METHOD get_stTankLevel : ST_Tank_Level
VAR_INPUT
END_VAR
VAR
	blank: ST_Tank_Level;
END_VAR
IF __ISVALIDREF(stTankLevel) THEN;
	get_stTankLevel:=stTankLevel;
ELSE;
	get_stTankLevel:=blank;
END_IF
END_METHOD

METHOD get_stTankLevel_OverFlow : BOOL
VAR_INPUT
END_VAR
VAR
	blank: ST_Tank_Level;
END_VAR
IF __ISVALIDREF(stTankLevel) THEN;
	IF stTankLevel.bIn_HL_signal 
	OR stTankLevel.rTankLevelPercentage>100
	OR (NOT MAIN.bTemp_Water_Overweight_check)
	THEN;
		get_stTankLevel_OverFlow:=TRUE;
	ELSE;
		get_stTankLevel_OverFlow:=FALSE;
	END_IF	
ELSE;
	get_stTankLevel_OverFlow:=FALSE;
END_IF
END_METHOD

END_FUNCTION_BLOCK

// ---- 00 Library/04 Recipe/FB_Recipe.TcPOU
FUNCTION_BLOCK FB_Recipe
VAR_INPUT
	pstRecipe				:POINTER TO ST_Recipe;
	bMemoRecipeUpdated		:BOOL:=FALSE;
	sRecipeDef				:STRING; (* current recipe definition *)
	bLoadDefault			:BOOL;
	sRecipesStoragePath		:STRING;
	bHMI_FrameActive		:BOOL;

END_VAR

VAR
	i						:INT;	
	RecipeManCommands 		:RecipeManCommands; (* Recipe Manager *)
	k						:INT;
	t1						:TON;
	check					:DWORD;
	INDEX					:INT:= 0;
	bReloadRecipes			:BOOL;
	rt_LoadDefault: R_TRIG;
	MessageBox			:MessageBox_Struct;
	arrLastReturn		: ARRAY[0..15] OF DWORD;
	LastReturn			:  DWORD;
	ton_RecipeUpdated: TON;
	sMessage: STRING;
	ton_SetStoragePath_Delay: TON;
	bSetStoragePath: BOOL:=TRUE;
	ton_SetStoragePathTimeOut: TON;
	bReturn: BOOL;
	
	ton_MessClear: TON;
	rt_Init: R_TRIG;
	sLastMessage: STRING;
	rt_Saved: R_TRIG;
	rt_FrameAvtive: R_TRIG;
	rt_LoadDefault1: R_TRIG;
END_VAR

act_SetStoragePath();
act_Disp();

IF pstRecipe^.bValidSelected THEN
	pstRecipe^.sSelectedReceipe:= pstRecipe^.arrRecipeNames[pstRecipe^.iRecipeIndex];
	pstRecipe^.bValidSelected:=FALSE;
END_IF

rt_FrameAvtive(CLK:=bHMI_FrameActive);
rt_LoadDefault1(CLK:=bLoadDefault);
IF pstRecipe^.bReInit OR rt_LoadDefault1.Q OR rt_FrameAvtive.Q THEN;
	pstRecipe^.bReInit:=FALSE;
	pstRecipe^.bInit:=FALSE;
	bSetStoragePath:=TRUE;
END_IF

t1(IN:=NOT pstRecipe^.bInit , PT:=T#0.5S);
IF (NOT pstRecipe^.bInit AND t1.Q) THEN
	
	IF NOT bSetStoragePath THEN;
		arrLastReturn[3]:=RecipeManCommands.ResetLastInfo();
		arrLastReturn[4]:=RecipeManCommands.ReloadRecipes(RecipeDefinitionName:=sRecipeDef);
		pstRecipe^.iRecipeCount:=RecipeManCommands.GetRecipeCount(sRecipeDef);
		FOR i := 0 TO GVL_Recipe.C_Max_RecipeFileNum DO
			pstRecipe^.arrRecipeNames[i] := '';
		END_FOR
		FOR i := 0 TO 1200 DO
			pstRecipe^.arrVariableNamesValue[i] := '';
			pstRecipe^.arrVariableValue[i] := '';
		END_FOR	
		(* save all recipe names of one recipe definition in an array *)
		arrLastReturn[0]:=RecipeManCommands.GetRecipeNames(sRecipeDef, ADR(pstRecipe^.arrRecipeNames),GVL_Recipe.C_Max_RecipeFileNum, 0);
		pstRecipe^.iRecipeIndex:=0;
		pstRecipe^.sLastSelectedReceipe:=pstRecipe^.sSelectedReceipe:=pstRecipe^.arrRecipeNames[0];
		pstRecipe^.bInit:=TRUE;
		pstRecipe^.bReInit:=FALSE;		
	END_IF

END_IF


rt_Init(CLK:=pstRecipe^.bInit);
IF pstRecipe^.bInit THEN

	IF pstRecipe^.sSelectedReceipe <> pstRecipe^.sLastSelectedReceipe 
	OR rt_Init.Q 
	OR rt_Saved.Q
	THEN;
				 
		arrLastReturn[1]:=RecipeManCommands.GetRecipeValues
			(
			RecipeDefinitionName:= sRecipeDef,
			RecipeName:= pstRecipe^.sSelectedReceipe, 
			pStrings:= ADR(pstRecipe^.arrVariableValue), 
			iSize:= 1200, 
			iStartIndex:= 0, 
			iStringLength:=80
			 );		
					
		arrLastReturn[2]:=RecipeManCommands.GetRecipeVariableNames
			(
			RecipeDefinitionName:=sRecipeDef,
			RecipeName:=pstRecipe^.sSelectedReceipe, 
			pStrings:= ADR(pstRecipe^.arrVariableNamesValue), 
			iSize:= 1200, 
			iStartIndex:= 0
			);
				
			pstRecipe^.bShowFile:=FALSE;
	END_IF
	pstRecipe^.sLastSelectedReceipe:=pstRecipe^.sSelectedReceipe;
END_IF


FOR i:=0 TO 15 DO
	IF arrLastReturn[i]<>0 THEN
		LastReturn:=arrLastReturn[i];
		EXIT;
	END_IF
	IF i=15 AND arrLastReturn[i]=0 THEN
		LastReturn:=0;
	END_IF
END_FOR

act_Cmd_List();

ACTION act_Cmd_List:
rt_LoadDefault(CLK:=bLoadDefault AND NOT bSetStoragePath);
IF rt_LoadDefault.Q THEN;
	pstRecipe^.sSelectedReceipe:='Default';
	pstRecipe^.bWriteToPLC_Cmd:=TRUE;
END_IF


IF pstRecipe^.bReloadRecipes THEN
	arrLastReturn[3]:=RecipeManCommands.ResetLastInfo();
	arrLastReturn[4]:=RecipeManCommands.ReloadRecipes(RecipeDefinitionName:=sRecipeDef);
	pstRecipe^.bReloadRecipes:=FALSE;
END_IF


IF pstRecipe^.bGetLastError THEN
	arrLastReturn[5]:=RecipeManCommands.GetLastError();
	pstRecipe^.bGetLastError:=FALSE;
END_IF


IF pstRecipe^.bResetLastError THEN
	arrLastReturn[6]:=RecipeManCommands.ResetLastError();
	pstRecipe^.bResetLastError:=FALSE;
	sMessage:='';
	FOR i:=0 TO 15 DO
		arrLastReturn[i]:=0;
	END_FOR	
END_IF

rt_Saved(CLK:=NOT pstRecipe^.bSaveFileCmd);
IF pstRecipe^.bSaveFileCmd  THEN
	sMessage:='cmd Save Recipe';
	IF  METH_Search(pstRecipe:=pstRecipe , sSearchRecipe:=pstRecipe^.sSelectedReceipe ) THEN
		//arrLastReturn[7]:=RecipeManCommands.ReadAndSaveRecipeAs(RecipeDefinitionName:=sRecipeDef,
		arrLastReturn[7]:=RecipeManCommands.ReadAndSaveRecipe(RecipeDefinitionName:=sRecipeDef,
			RecipeName:=pstRecipe^.sSelectedReceipe);// ,
			//FileName:='.txtrecipe' );
		sMessage:='cmd Save Recipe - Done';
		pstRecipe^.bSaveFileCmd:=FALSE;
	ELSE;
		sMessage:='cmd Save Recipe - Failed';
	END_IF
END_IF


IF pstRecipe^.bWriteToPLC_Cmd  THEN
	sMessage:='cmd Load Recipe';
	bMemoRecipeUpdated:=FALSE;
	IF  METH_Search(pstRecipe:=pstRecipe , sSearchRecipe:=pstRecipe^.sSelectedReceipe ) THEN
		arrLastReturn[8]:=RecipeManCommands.LoadRecipe(RecipeDefinitionName:= sRecipeDef, RecipeName:= pstRecipe^.sSelectedReceipe);
		arrLastReturn[9]:=RecipeManCommands.WriteRecipe(RecipeDefinitionName:= sRecipeDef, RecipeName:= pstRecipe^.sSelectedReceipe);
		sMessage:='cmd Load Recipe - Done';
		pstRecipe^.bWriteToPLC_Cmd:=FALSE;
		ton_RecipeUpdated.IN:=TRUE;
	ELSE;
		sMessage:='cmd Load Recipe - Failed';
	END_IF
END_IF
ton_RecipeUpdated(PT:=T#1S);
IF ton_RecipeUpdated.Q THEN;
	bMemoRecipeUpdated:=TRUE;	
	ton_RecipeUpdated.IN:=FALSE;
END_IF


IF pstRecipe^.bCreateRecipe AND pstRecipe^.sNewRecipeName <> '' THEN
	arrLastReturn[10]:=RecipeManCommands.CreateRecipe(sRecipeDef ,pstRecipe^.sNewRecipeName);
	sMessage:='cmd Create Recipe - Done';
	pstRecipe^.bCreateRecipe:=FALSE;
	pstRecipe^.bReInit:=TRUE;
END_IF


IF pstRecipe^.bDeleteRecipe THEN
	sMessage:='cmd Delete Recipe';
	IF  METH_Search(pstRecipe:=pstRecipe , sSearchRecipe:=pstRecipe^.sSelectedReceipe ) THEN
		arrLastReturn[11]:=RecipeManCommands.DeleteRecipe(sRecipeDef ,pstRecipe^.sSelectedReceipe);
		sMessage:='cmd Delete Recipe - Done';
		pstRecipe^.bDeleteRecipe:=FALSE;
		pstRecipe^.bReInit:=TRUE;
	ELSE;
		sMessage:='cmd Delete Recipe - Failed';
	END_IF
END_IF

ton_MessClear(PT:=T#30S);
IF sMessage<>sLastMessage THEN;
	ton_MessClear(IN:=FALSE);
	sLastMessage:=sMessage;
ELSIF sMessage<>'' THEN;
	ton_MessClear.IN:=TRUE;
ELSE;
	ton_MessClear.IN:=FALSE;
END_IF
IF ton_MessClear.Q THEN;
	sMessage:='';
END_IF
END_ACTION

ACTION act_Disp:

IF pstRecipe^.iDispSel<0 THEN; pstRecipe^.iDispSel:=0; END_IF
IF pstRecipe^.iDispSel>1180 THEN; pstRecipe^.iDispSel:=1180; END_IF

//FOR k:=iDispSel TO iDispSel+19 DO;
FOR k:=0 TO 20 DO;
	pstRecipe^.arrVariableDisp[0,k]:= INT_TO_STRING(pstRecipe^.iDispSel+k);
	pstRecipe^.arrVariableDisp[1,k]:=pstRecipe^.arrVariableNamesValue[pstRecipe^.iDispSel+k];
	pstRecipe^.arrVariableDisp[2,k]:=pstRecipe^.arrVariableValue[pstRecipe^.iDispSel+k];
END_FOR
END_ACTION

ACTION act_SetStoragePath:
ton_SetStoragePath_Delay(PT:=T#0.5S,IN:=bSetStoragePath);
ton_SetStoragePathTimeOut(PT:=T#2S);

IF ton_SetStoragePath_Delay.Q THEN;
	bReturn:=RecipeManCommands.SetStoragePath(stPath:=sRecipesStoragePath);
	//sMessage:='cmd Set Storage Path';
	IF bReturn THEN;
		bSetStoragePath:=FALSE;
		ton_SetStoragePathTimeOut.IN:=FALSE;
		//sMessage:='cmd Set Storage Path - Done';
	ELSE
		ton_SetStoragePathTimeOut.IN:=TRUE;
	END_IF
	
	IF ton_SetStoragePathTimeOut.Q THEN;
		bSetStoragePath:=FALSE;
		ton_SetStoragePathTimeOut.IN:=FALSE;
		//sMessage:='cmd Set Storage Path - Failed';		
	END_IF
END_IF
END_ACTION

METHOD METH_Search : BOOL
VAR_INPUT
	pstRecipe :POINTER TO ST_Recipe;
	sSearchRecipe	:STRING(30);
END_VAR

VAR
	i: INT;
END_VAR
METH_Search:=FALSE;
FOR i:= 0 TO GVL_Recipe.C_Max_RecipeFileNum DO
	IF sSearchRecipe = pstRecipe^.arrRecipeNames[i] THEN
		METH_Search:=TRUE;
		EXIT;
	END_IF
END_FOR
END_METHOD

END_FUNCTION_BLOCK

// ---- 00 Library/04-Messages/FB_PrintErrMessageByID.TcPOU
FUNCTION_BLOCK FB_PrintErrMessageByID
VAR_INPUT
	sActErrorID			: STRING;
	iFB_Num				: INT:=0;
	sModuleDescription	:STRING:='';
END_VAR
VAR_OUTPUT
END_VAR
VAR
	cFound				: INT;
	i					: INT;
	iFound				: INT;
	bNewMeasege			: BOOL;
	rtrig1				: R_TRIG;
	sLastErrorID		: STRING;
	j: INT;
	sFB_Num: STRING(3);

END_VAR




	
	IF sActErrorID<>'000x000x000'  AND sActErrorID<>'' THEN
		IF iFB_Num>0 THEN;
			sFB_Num:=F_iFB_Num_sFB_Num(iFB_Num:=iFB_Num);
			sLastErrorID:=REPLACE(sActErrorID,sFB_Num,3,5);
		ELSE;
			sLastErrorID:=sActErrorID;
		END_IF			
		
		bNewMeasege:=TRUE;
		FOR i:=1 TO 100 DO
			IF Buffer_Act_Message[i].sErrID=sLastErrorID THEN;//sActErrorID
				//IF Buffer_Act_Message[i].sModuleDescription = sFB_ModuleDescription THEN
					bNewMeasege:=FALSE;
					EXIT; 
				//END_IF
			END_IF
		END_FOR
	ELSE
		bNewMeasege:=FALSE;
	END_IF
	
	IF bNewMeasege THEN;
		FOR i:=100 TO 2 BY -1 DO
			Buffer_Act_Message[i].sDateTime:=Buffer_Act_Message[i-1].sDateTime;
			Buffer_Act_Message[i].sErrID:=Buffer_Act_Message[i-1].sErrID;
			Buffer_Act_Message[i].sErrorMessage:=Buffer_Act_Message[i-1].sErrorMessage;
			Buffer_Act_Message[i].sLevel:=Buffer_Act_Message[i-1].sLevel;
			Buffer_Act_Message[i].sModuleDescription:=Buffer_Act_Message[i-1].sModuleDescription;
		END_FOR
		
		Buffer_Act_Message[1].sDateTime:=prg_RealClock.sRealTime_Date;
		Buffer_Act_Message[1].sErrID:=sLastErrorID;//sActErrorID
		Buffer_Act_Message[1].sModuleDescription:=sModuleDescription;

		//IF sActErrorID='000x000x999' THEN;
		//	Buffer_Act_Message[1].sErrorMessage:='General Error';	(*	Error description Not Found	*)
		//ELSE
			cFound:=0;
			FOR i:=1 TO C_Max_ErrorList DO
				IF ar_ErrorList[i,eErrID]=sActErrorID THEN
					iFound:=i;
					ar_ErrorActive[iFound]:=TRUE;
					cFound:=cFound+1;
				END_IF
			END_FOR
	
			IF cFound=1 THEN;
				Buffer_Act_Message[1].sErrorMessage:=ar_ErrorList[iFound,eErrMeassage];	(*	Error from the List	*)
				Buffer_Act_Message[1].sLevel:=ar_ErrorList[iFound,eErrLevel];	(*	Error Level from the List	*)
			ELSIF cFound=0 THEN; //(*	Error ID not Foud on the Error_List*)
				Buffer_Act_Message[1].sErrorMessage:='Error ID not found on the "Error_List"';	
				Buffer_Act_Message[1].sLevel:='Unknown';
			ELSIF cFound>1 THEN; //(*	More then one Errors Foud with the same  ID*)
				Buffer_Act_Message[1].sErrorMessage:='More then one error with the same ID  found on the "Error_list"';	
				Buffer_Act_Message[1].sLevel:='Unknown';
			END_IF
		//END_IF
		FUN_Write_Line_To_History();
	END_IF

END_FUNCTION_BLOCK

// ---- 00 Library/04-Messages/F_iFB_Num_sFB_Num.TcPOU
FUNCTION F_iFB_Num_sFB_Num : STRING(3)
VAR_INPUT
	iFB_Num: INT;
END_VAR
VAR
END_VAR

IF iFB_Num<10 THEN;
	F_iFB_Num_sFB_Num:=CONCAT(STR1:='00',STR2:=INT_TO_STRING(iFB_Num));
ELSIF iFB_Num<100 THEN;
	F_iFB_Num_sFB_Num:=CONCAT(STR1:='0',STR2:=INT_TO_STRING(iFB_Num));
ELSE;
	F_iFB_Num_sFB_Num:=CONCAT(STR1:='',STR2:=INT_TO_STRING(iFB_Num));
END_IF

END_FUNCTION

// ---- 00 Library/03 SFC/FB_SFC_Template.TcPOU
FUNCTION_BLOCK FB_SFC_Template EXTENDS FB_SFC_Cycle IMPLEMENTS ITF_FB_SFC_Cycle
VAR_INPUT
END_VAR
VAR_OUTPUT
END_VAR
VAR
END_VAR

m_Set_SFCFlags_Reference();
SUPER^();

ACTION act_Oper:
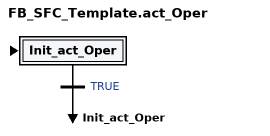
INITIAL_STEP Init_act_Oper:
END_STEP
TRANSITION FROM Init_act_Oper TO Init_act_Oper
    := TRUE;
END_TRANSITION
END_ACTION

METHOD m_Set_SFCFlags_Reference : BOOL
//Set reference to SFC flags

refSFC.SFCInit REF= SFCInit;
refSFC.SFCReset REF= SFCReset;
refSFC.SFCError REF= SFCError;
refSFC.SFCEnableLimit REF= SFCEnableLimit;
refSFC.SFCErrorStep REF= SFCErrorStep;
refSFC.SFCErrorPOU REF= SFCErrorPOU;
refSFC.SFCQuitError REF= SFCQuitError;
refSFC.SFCPause REF= SFCPause;
refSFC.SFCTrans REF= SFCTrans;
refSFC.SFCCurrentStep REF= SFCCurrentStep;
refSFC.SFCTip REF= SFCTip;
refSFC.SFCTipMode REF= SFCTipMode;

// Cycle handle for SFC
m_SFC_Handle();
END_METHOD

END_FUNCTION_BLOCK

// ---- 03 Project/00 -Initialise/prg_Initialise.TcPOU
PROGRAM prg_Initialise
VAR_INPUT
	ResumeSFC       : BOOL; 		(*	not automatic	*)
	//Added SFC Cycle handle Variables
	
	SFCInit             : BOOL;  //shachar
END_VAR

VAR


(* 8888888888888888   SFC   8888888888888888888888*)
	sCycleName	        : STRING;
	SFCCurrentStep      : STRING;
	SFCErrorPOU         : STRING;
	SFCErrorStep        : STRING;
	SFCError            : BOOL;
	SFCPause            : BOOL;
	
	SFCTipMode          : BOOL;
	SFCTip              : BOOL;
	SFCEnableLimit		: BOOL:=TRUE;
	// Reset Error
	SFCReset			: BOOL;
	ErrorSFC            : BOOL; 	(*	not automatic	*)

	ResetError          : BOOL; 	(*	not automatic	*)
	Last_SFCErrorStep   : STRING; 	(*	not automatic	*)
	//ErrorToPrint        : STRING; 	(*	not automatic	*)
	//Last_ErrorToPrint   : STRING; 	(*	not automatic	*)

 //   stSafety			:ST_BasicCycle;  //shachar
(* 8888888888888888   SFC   8888888888888888888888*)




	Pis             : INT;
	c_PisInitCheck  : INT;
	b_AllPisInitPos : BOOL;

	i               : INT;
	c_LatInitCheck  : INT;

	c_PisResetCleare: INT;

	k               : INT;

	bGeneralDone    : BOOL;
	bPistonDone     : BOOL;
	b_StationDone   : BOOL;
	bLoadConvDone   : BOOL;
	bUnloadConvDone : BOOL;
	bTableDone      : BOOL;
	bStackerDone    : BOOL;
    bManipulatorDone: BOOL;

	init_General    : BOOL;
	init_AllPiston  : BOOL;
	init_AllStation : BOOL;
	init_Table      : BOOL;
	init_LoadConv   : BOOL;
	init_UnloadConv : BOOL;
	init_Stacker    : BOOL;
	init_Manipulator: BOOL;

	bMessLoadInit   : BOOL;
	bMessUnloadInit : BOOL;
	
	sFB_ID          : STRING(4):='004';
	sFB_Num         : STRING(4):='000';
	sActErrorID     : STRING;
	//Added SFC Cycle handle Variables
	fb_SFC_Cycle		    : FB_SFC_Cycle;
	fbFormatString	    	: FB_FORMATSTRING;
	sFullErrorId		    : STRING(12);//sAAAxBBBxEEE
	bReset					: BOOL;

	bIntZoneOk: BOOL;
	bNotPrepare: BOOL;
	p_ManipReset: POINTER TO BOOL;
	p_PowerMotorOn: POINTER TO BOOL;
	p_SafetyStart: POINTER TO BOOL;
   // fbPowerMotorOn			:FB_PowerMotorOn;

	IndexOn: BOOL;
	LoadOn: BOOL;
	UnloadOn: BOOL;
	ManipOn: BOOL;
	p_PowerMotorPower: POINTER TO BOOL;
	p_PowerMotorOff: POINTER TO BOOL;
	iResumeCount: INT;
	iIndexCount: INT;
	iLoadCount: INT;
	iUnloadCount: INT;
	iManipCount: INT;
	p_ManipResume: POINTER TO BOOL;
END_VAR

VAR_IN_OUT
	stOperation	: ST_OperationButtons;	
END_VAR

act_General();
act_Piston();
act_GetErrorID();
fb_SFC_Cycle
( 
	sCycleName:= 'Initialize', 
	bSFCError:= SFCError, 
	sSFCCurrentStep:=SFCCurrentStep , 
	sSFCErrorStep:= SFCErrorStep, 
	sSFCErrorPOU:=SFCErrorPOU , 
	sActErrorID:=sFullErrorId,
	sFB_ModuleDescription:= fb_SFC_Cycle.sCycleName, 
	sLast_SFCErrorStep=>Last_SFCErrorStep , 
	bErrorSFC_Occured=> ErrorSFC, 
	//sErrorToPrint=>ErrorToPrint , 
	//sLast_ErrorToPrint=>Last_ErrorToPrint,
    bSFCInit=>SFCInit , 
	stOperation:= stOperation,
	bResumeSFC:=ResumeSFC , 
	bResetError:=ResetError , 
	bSFCPause:= SFCPause, 
	bResetCycle:=SFCReset
);



IF NOT bStateSafe	
OR init_AllPiston
THEN;
	bGeneralDone:=FALSE;
	bPistonDone:=FALSE;
	b_StationDone:=FALSE;
	bLoadConvDone:=FALSE;
	bUnloadConvDone:=FALSE;
	bTableDone:=FALSE;
	bStackerDone:=FALSE;
	bManipulatorDone:=FALSE;  //shachar
END_IF

ACTION act_General:
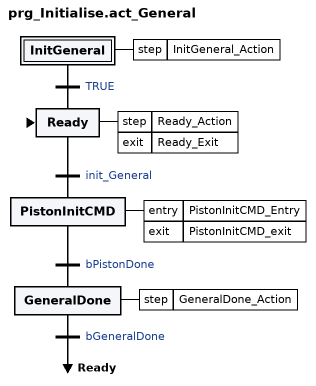
INITIAL_STEP InitGeneral:
    InitGeneral_Action(N);  // step action
END_STEP
TRANSITION FROM InitGeneral TO Ready
    := TRUE;
END_TRANSITION
STEP Ready:
    Ready_Action(N);  // step action
    Ready_Exit(P0);  // exit action
END_STEP
TRANSITION FROM Ready TO PistonInitCMD
    := init_General;
END_TRANSITION
STEP PistonInitCMD:  // min time t#2s
    PistonInitCMD_Entry(P1);  // entry action
    PistonInitCMD_exit(P0);  // exit action
END_STEP
TRANSITION FROM PistonInitCMD TO GeneralDone
    := bPistonDone;
END_TRANSITION
STEP GeneralDone:
    GeneralDone_Action(N);  // step action
END_STEP
TRANSITION FROM GeneralDone TO Ready
    := bGeneralDone;
END_TRANSITION
END_ACTION

ACTION act_GetErrorID:
IF ErrorSFC THEN;
	// Initialization
	IF    Last_SFCErrorStep='WatingForEmergencyOK' 			THEN sActErrorID:='001';
	ELSIF Last_SFCErrorStep='WatingForInterlockOK' 		    THEN sActErrorID:='002';
	ELSIF Last_SFCErrorStep='WatingForMotorsOK' 			THEN sActErrorID:='003';
	ELSIF Last_SFCErrorStep='CheckInitStationDone' 			THEN sActErrorID:='004';
	ELSIF Last_SFCErrorStep='Station_Initialization' 		THEN sActErrorID:='005';
	ELSIF Last_SFCErrorStep='Loader_Initialization' 		THEN sActErrorID:='006';
	ELSIF Last_SFCErrorStep='Unload_Station' 			    THEN sActErrorID:='007';
	ELSIF Last_SFCErrorStep='Measuring_Station' 			THEN sActErrorID:='008';
	ELSIF Last_SFCErrorStep='Gripper_Oriantation' 			THEN sActErrorID:='009';
	ELSIF Last_SFCErrorStep='Index_Homming' 			    THEN sActErrorID:='010';
	ELSIF Last_SFCErrorStep='PaletBypasCheck_1' 			THEN sActErrorID:='011';
	ELSIF Last_SFCErrorStep='PaletCheck_1' 			        THEN sActErrorID:='012';
	ELSIF Last_SFCErrorStep='Cover_Station' 			    THEN sActErrorID:='023';	
	ELSE;
		 sActErrorID:='999';
	END_IF
//ELSIF bWarning THEN;
	// Leave the warning message to print
ELSE;
		 sActErrorID:='000';
END_IF
//*** Error Format ***
fbFormatString(
	sFormat:= '%.3sx%.3sx%.3s', 
	arg1:= F_STRINGEx(sFB_ID), 
	arg2:= F_STRINGEx(sFB_Num), 
	arg3:= F_STRINGEx(sActErrorID), 
	sOut=>sFullErrorId );
	
//(*Clean Last ErrID*)IF NOT SFCPause THEN	sFullErrorId:='';END_IF
END_ACTION

ACTION act_Piston:
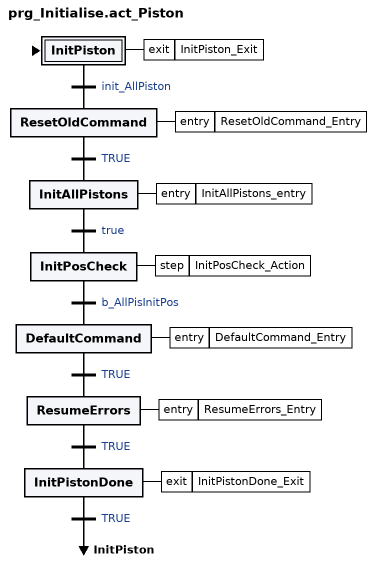
INITIAL_STEP InitPiston:
    InitPiston_Exit(P0);  // exit action
END_STEP
TRANSITION FROM InitPiston TO ResetOldCommand
    := init_AllPiston;
END_TRANSITION
STEP ResetOldCommand:  // min time T#0.1S
    ResetOldCommand_Entry(P1);  // entry action
END_STEP
TRANSITION FROM ResetOldCommand TO InitAllPistons
    := TRUE;
END_TRANSITION
STEP InitAllPistons:  // min time t#1s
    InitAllPistons_entry(P1);  // entry action
END_STEP
TRANSITION FROM InitAllPistons TO InitPosCheck
    := true;
END_TRANSITION
STEP InitPosCheck:
    InitPosCheck_Action(N);  // step action
END_STEP
TRANSITION FROM InitPosCheck TO DefaultCommand
    := b_AllPisInitPos;
END_TRANSITION
STEP DefaultCommand:  // min time T#0.2S
    DefaultCommand_Entry(P1);  // entry action
END_STEP
TRANSITION FROM DefaultCommand TO ResumeErrors
    := TRUE;
END_TRANSITION
STEP ResumeErrors:  // min time T#0.2S
    ResumeErrors_Entry(P1);  // entry action
END_STEP
TRANSITION FROM ResumeErrors TO InitPistonDone
    := TRUE;
END_TRANSITION
STEP InitPistonDone:
    InitPistonDone_Exit(P0);  // exit action
END_STEP
TRANSITION FROM InitPistonDone TO InitPiston
    := TRUE;
END_TRANSITION
END_ACTION

ACTION DefaultCommand_Entry:
	(*FOR Pis:=1 TO 24 BY 1 DO
		db_Lat[Pis].req_DefaultPos:=TRUE;
	END_FOR*)
	
	FOR Pis:=1 TO C_Max_Pistons BY 1 DO
		IF stPis[Pis].b_PistonActive THEN;
			stPis[Pis].req_Init:=TRUE;
		END_IF		
	END_FOR
END_ACTION

ACTION GeneralDone_Action:
init_General:=FALSE;
bGeneralDone:=TRUE;
END_ACTION

ACTION InitAllPistons_entry:
prg_Pistons.bInitAllPiston:=TRUE;
END_ACTION

ACTION InitGeneral_Action:
SFCReset:=FALSE;

init_AllPiston   :=FALSE;
END_ACTION

ACTION InitPiston_Exit:
	b_AllPisInitPos:=FALSE;
	bPistonDone:=FALSE;
END_ACTION

ACTION InitPistonDone_Exit:
	init_AllPiston:=FALSE;
	bPistonDone:=TRUE;
END_ACTION

ACTION InitPosCheck_Action:
			c_PisInitCheck:=0;
	FOR Pis:=1 TO C_Max_Pistons BY 1 DO
		IF fb_Pis[Pis].SFCCurrentStep<>'Ready' AND fb_Pis[Pis].SFCCurrentStep<>''THEN
			c_PisInitCheck:=c_PisInitCheck+1;
		END_IF
	END_FOR

			c_PisResetCleare:=0;
	FOR Pis:=1 TO C_Max_Pistons BY 1 DO
		IF stPis[Pis].b_Reset THEN
			c_PisResetCleare:=c_PisResetCleare+1;
		END_IF
	END_FOR

	(*		c_LatInitCheck:=0;
	FOR Pis:=1 TO 24 BY 1 DO
		IF fb_Lat[Pis].SFCCurrentStep<>'Ready' AND fb_Lat[Pis].SFCCurrentStep<>'' THEN
			c_LatInitCheck:=c_LatInitCheck+1;
		END_IF
	END_FOR*)


		IF 	c_PisInitCheck=0  AND c_LatInitCheck=0 (*AND 	c_PisResetCleare=0*) THEN
			b_AllPisInitPos:=TRUE;
		ELSE
			b_AllPisInitPos:=FALSE;
		END_IF
END_ACTION

ACTION PistonInitCMD_Entry:
init_AllPiston:=TRUE;
END_ACTION

ACTION PistonInitCMD_exit:
Global_Variables.ResumeAll :=TRUE;
END_ACTION

ACTION Ready_Action:
IF TRUE
AND	bPistonDone
(*AND	b_StationDone
AND	bLoadConvDone
AND	bUnloadConvDone
AND	bTableDone
AND (bManipulatorDone OR NOT b_ManipulatorExist)
AND	(bStackerDone OR NOT b_StackerExist)*)
THEN
	bGeneralDone:=TRUE;

ELSE
	bGeneralDone:=FALSE;
END_IF
END_ACTION

ACTION Ready_Exit:
bGeneralDone:=FALSE;
bPistonDone:=FALSE;
b_StationDone:=FALSE;
bLoadConvDone:=FALSE;
bUnloadConvDone:=FALSE;
bTableDone:=FALSE;
bStackerDone:=FALSE;

bManipulatorDone:=FALSE; //shachar
iResumeCount:=0;
END_ACTION

ACTION ResetOldCommand_Entry:
	(*FOR Pis:=1 TO 24 BY 1 DO
		db_Lat[Pis].req_Reset:=TRUE;
	END_FOR*)
	FOR Pis:=1 TO C_Max_Pistons BY 1 DO
		stPis[Pis].b_Reset:=TRUE;
	END_FOR
END_ACTION

ACTION ResumeErrors_Entry:
	(*FOR Pis:=1 TO 24 BY 1 DO
		db_Lat[Pis].req_Resume:=TRUE;
	END_FOR*)
	FOR Pis:=1 TO C_Max_Pistons BY 1 DO
		stPis[Pis].b_Resume:=TRUE;
	END_FOR
END_ACTION

END_PROGRAM

// ---- 03 Project/31 AnybusCommunication/FB_Anybus_Interface.TcPOU
//CIP <-> Siemens exchange through the Anybus Communicator, 128 bytes each direction.
//Spec: "Интерфейс CIP ↔ Siemens через Anybus", meeting 28.10.2026.
//Decodes the Siemens data, checks ALIVE and the values, encodes the CIP status.
//While communication is lost all Siemens inputs are treated as 0 (REQUEST ON drops -> CIP pause).
FUNCTION_BLOCK FB_Anybus_Interface
VAR_INPUT
	stStatus		: ST_Anybus_Outputs;	//CIP -> Siemens, filled by the CIP logic (bAlive is generated here)
	bFieldbusOk		: BOOL := TRUE;			//gateway EtherCAT slave: WcState = 0 (gIO.Anybus_WcState in MAIN)
	bSwapBytes		: BOOL := TRUE;			//TRUE: INT/DINT are big-endian (Profinet), swapped here
	tAliveTimeout	: TIME := T#2S;			//Siemens ALIVE must toggle within this time
	tNextStable		: TIME := T#3S;			//NEXT CLIENT / NEXT RECIPE must be stable this long
END_VAR
VAR_IN_OUT
	arRawIn			: ARRAY[0..127] OF BYTE;	//gIO.Anybus_Inputs_Raw
	arRawOut		: ARRAY[0..127] OF BYTE;	//gIO.Anybus_Outputs_Raw
END_VAR
VAR_OUTPUT
	stIn			: ST_Anybus_Inputs;		//Siemens -> CIP, all 0 while communication is lost
	stOut			: ST_Anybus_Outputs;	//CIP -> Siemens as actually sent (with ALIVE, alarm bit and code)
	bCommOk			: BOOL;					//fieldbus OK and Siemens ALIVE toggles
	eRequest		: E_Anybus_Request;		//combination of REQUEST ON / REQUEST OFF
	bRequestOnEdge	: BOOL;					//one cycle when eRequest becomes eOn (start or resume)
	bRequestOffEdge	: BOOL;					//one cycle when eRequest becomes eOff
	bCurrentValid	: BOOL;					//CLIENT ID, RECIPE TYPE, CLIENT TYPE are in range
	bNextValid		: BOOL;					//next client is in range and stable for tNextStable
	nNextClient		: INT;					//accepted next client, 0 = none
	eNextRecipe		: E_Anybus_RecipeType;	//accepted next recipe
	eNextClientType	: E_Anybus_ClientType;	//accepted next client type, eNone = not sent
	eAlarm			: E_Anybus_Alarm;		//interface alarm, eNone = OK
END_VAR
VAR
	stRaw			: ST_Anybus_Inputs;		//decoded, before the communication check
	stBlank			: ST_Anybus_Inputs;

	//ALIVE
	bAliveOut		: BOOL;
	tonAliveOut		: TON;
	tonAliveIn		: TON;
	bAliveInMemo	: BOOL;
	bAliveSeen		: BOOL;					//at least one toggle since start

	rtRequestOn		: R_TRIG;
	rtRequestOff	: R_TRIG;

	//Next client
	tonNextStable	: TON;
	nNextClientMemo	: INT;
	eNextRecipeMemo	: E_Anybus_RecipeType;
	eNextTypeMemo	: E_Anybus_ClientType;
	bNextInRange	: BOOL;
END_VAR
VAR CONSTANT
	cnClientMax		: INT := 30;
END_VAR

//Decode Siemens -> CIP
//Bits are addressed by byte (Siemens x.y = byte x, bit y), no swap
stRaw.bAlarm			:= arRawIn[0].0;
stRaw.bReady			:= arRawIn[0].1;
stRaw.bRequestOn		:= arRawIn[0].2;
stRaw.bRequestOff		:= arRawIn[0].3;
stRaw.bInletPumpEnable	:= arRawIn[0].4;
stRaw.bPause			:= arRawIn[0].5;
stRaw.bClientEmpty		:= arRawIn[0].6;
stRaw.bAlive			:= arRawIn[0].7;
stRaw.bSprinklerState	:= arRawIn[1].0;
stRaw.nClientId			:= m_GetInt(arRaw:=arRawIn, nWord:=1);
stRaw.eRecipeType		:= m_GetInt(arRaw:=arRawIn, nWord:=2);
stRaw.eClientType		:= m_GetInt(arRaw:=arRawIn, nWord:=3);
stRaw.nNextClient		:= m_GetInt(arRaw:=arRawIn, nWord:=4);
stRaw.eNextRecipe		:= m_GetInt(arRaw:=arRawIn, nWord:=5);
stRaw.eNextClientType	:= m_GetInt(arRaw:=arRawIn, nWord:=6);

//Siemens ALIVE watchdog
IF stRaw.bAlive <> bAliveInMemo THEN;
	bAliveInMemo:=stRaw.bAlive;
	bAliveSeen:=TRUE;
	tonAliveIn(IN:=FALSE);
END_IF
tonAliveIn(IN:=TRUE, PT:=tAliveTimeout);
bCommOk:=bFieldbusOk AND bAliveSeen AND NOT tonAliveIn.Q;

//Communication lost: the same as the gateway clearing the data
IF bCommOk THEN;
	stIn:=stRaw;
ELSE;
	stIn:=stBlank;
END_IF

//REQUEST ON / REQUEST OFF
IF stIn.bRequestOn AND stIn.bRequestOff THEN;
	eRequest:=E_Anybus_Request.eConflict;
ELSIF stIn.bRequestOn THEN;
	eRequest:=E_Anybus_Request.eOn;
ELSIF stIn.bRequestOff THEN;
	eRequest:=E_Anybus_Request.eOff;
ELSE;
	eRequest:=E_Anybus_Request.eNone;
END_IF
rtRequestOn(CLK:=eRequest=E_Anybus_Request.eOn);
bRequestOnEdge:=rtRequestOn.Q;
rtRequestOff(CLK:=eRequest=E_Anybus_Request.eOff);
bRequestOffEdge:=rtRequestOff.Q;

//Current client: checked here, latched by the CIP logic on bRequestOnEdge
bCurrentValid:=TRUE
	AND stIn.nClientId>=1 AND stIn.nClientId<=cnClientMax
	AND stIn.eRecipeType>=E_Anybus_RecipeType.eFlushOnly AND stIn.eRecipeType<=E_Anybus_RecipeType.eFull
	AND stIn.eClientType>=E_Anybus_ClientType.ePipe AND stIn.eClientType<=E_Anybus_ClientType.eTank;

//Next client: any change cancels the accepted one, new values are taken after tNextStable
bNextInRange:=TRUE
	AND stIn.nNextClient>=1 AND stIn.nNextClient<=cnClientMax
	AND stIn.eNextRecipe>=E_Anybus_RecipeType.eFlushOnly AND stIn.eNextRecipe<=E_Anybus_RecipeType.eFull
	AND stIn.eNextClientType>=E_Anybus_ClientType.eNone AND stIn.eNextClientType<=E_Anybus_ClientType.eTank;
IF stIn.nNextClient<>nNextClientMemo
OR stIn.eNextRecipe<>eNextRecipeMemo
OR stIn.eNextClientType<>eNextTypeMemo
THEN;
	nNextClientMemo:=stIn.nNextClient;
	eNextRecipeMemo:=stIn.eNextRecipe;
	eNextTypeMemo:=stIn.eNextClientType;
	tonNextStable(IN:=FALSE);
	bNextValid:=FALSE;
	nNextClient:=0;
	eNextRecipe:=E_Anybus_RecipeType.eNone;
	eNextClientType:=E_Anybus_ClientType.eNone;
END_IF
tonNextStable(IN:=bNextInRange, PT:=tNextStable);
IF tonNextStable.Q AND NOT bNextValid THEN;
	bNextValid:=TRUE;
	nNextClient:=nNextClientMemo;
	eNextRecipe:=eNextRecipeMemo;
	eNextClientType:=eNextTypeMemo;
END_IF

//Interface alarm, first cause wins
IF NOT bFieldbusOk THEN;
	eAlarm:=E_Anybus_Alarm.eFieldbus;
ELSIF NOT bCommOk THEN;
	eAlarm:=E_Anybus_Alarm.eAliveLost;
ELSIF eRequest=E_Anybus_Request.eConflict THEN;
	eAlarm:=E_Anybus_Alarm.eRequestConflict;
ELSIF stIn.bRequestOn AND (stIn.nClientId<1 OR stIn.nClientId>cnClientMax) THEN;
	eAlarm:=E_Anybus_Alarm.eInvalidClient;
ELSIF stIn.bRequestOn AND NOT (stIn.eRecipeType>=E_Anybus_RecipeType.eFlushOnly AND stIn.eRecipeType<=E_Anybus_RecipeType.eFull) THEN;
	eAlarm:=E_Anybus_Alarm.eInvalidRecipe;
ELSIF stIn.bRequestOn AND NOT bCurrentValid THEN;
	eAlarm:=E_Anybus_Alarm.eInvalidClientType;
ELSE;
	eAlarm:=E_Anybus_Alarm.eNone;
END_IF

//CIP ALIVE, 0.5 s / 0.5 s
tonAliveOut(IN:=NOT tonAliveOut.Q, PT:=T#500MS);
IF tonAliveOut.Q THEN;
	bAliveOut:=NOT bAliveOut;
END_IF

//CIP -> Siemens as sent: ALIVE generated here, interface alarm added
stOut:=stStatus;
stOut.bAlive:=bAliveOut;
stOut.bAlarm:=stStatus.bAlarm OR (eAlarm<>E_Anybus_Alarm.eNone);
//CIP alarm code first, interface alarm code otherwise
IF stOut.nAlarmCode=0 THEN;
	stOut.nAlarmCode:=eAlarm;
END_IF

//Encode CIP -> Siemens
arRawOut[0].0	:= stOut.bAlarm;
arRawOut[0].1	:= stOut.bReady;
arRawOut[0].2	:= stOut.bWorking;
arRawOut[0].3	:= stOut.bFinish;
arRawOut[0].4	:= stOut.bEmptyingClient;
arRawOut[0].5	:= stOut.bSendingPump;
arRawOut[0].6	:= stOut.bPause;
arRawOut[0].7	:= stOut.bAlive;
arRawOut[1]		:= 0;
arRawOut[1].0	:= stOut.bSprinklerRequest;
m_SetInt(arRaw:=arRawOut, nWord:=1, nValue:=stOut.eActualMedia);
m_SetDint(arRaw:=arRawOut, nWord:=2, nValue:=stOut.nRecipeProgress);
m_SetDint(arRaw:=arRawOut, nWord:=4, nValue:=stOut.nActualProgress);
m_SetInt(arRaw:=arRawOut, nWord:=6, nValue:=stOut.nAlarmCode);
m_SetInt(arRaw:=arRawOut, nWord:=7, nValue:=stOut.nProgressUnit);
m_SetInt(arRaw:=arRawOut, nWord:=8, nValue:=stOut.nActiveClient);
m_SetInt(arRaw:=arRawOut, nWord:=9, nValue:=stOut.eActiveRecipe);
m_SetInt(arRaw:=arRawOut, nWord:=10, nValue:=stOut.nFlowRateSet);
m_SetInt(arRaw:=arRawOut, nWord:=11, nValue:=stOut.nFlowRateActual);

//INT of word nWord (bytes 2n, 2n+1)
METHOD PRIVATE m_GetInt : INT
VAR_IN_OUT
	arRaw	: ARRAY[0..127] OF BYTE;
END_VAR
VAR_INPUT
	nWord	: INT;
END_VAR
VAR
	nHi		: INT;	//byte index of the high byte
	nLo		: INT;	//byte index of the low byte
END_VAR
IF bSwapBytes THEN;
	nHi:=2*nWord;
	nLo:=2*nWord+1;
ELSE;
	nHi:=2*nWord+1;
	nLo:=2*nWord;
END_IF
m_GetInt:=WORD_TO_INT(SHL(BYTE_TO_WORD(arRaw[nHi]), 8) OR BYTE_TO_WORD(arRaw[nLo]));
END_METHOD

//Writes INT to word nWord (bytes 2n, 2n+1)
METHOD PRIVATE m_SetInt : BOOL
VAR_IN_OUT
	arRaw	: ARRAY[0..127] OF BYTE;
END_VAR
VAR_INPUT
	nWord	: INT;
	nValue	: INT;
END_VAR
VAR
	wValue	: WORD;
END_VAR
wValue:=INT_TO_WORD(nValue);
IF bSwapBytes THEN;
	arRaw[2*nWord]		:= WORD_TO_BYTE(SHR(wValue, 8));
	arRaw[2*nWord+1]	:= WORD_TO_BYTE(wValue);
ELSE;
	arRaw[2*nWord]		:= WORD_TO_BYTE(wValue);
	arRaw[2*nWord+1]	:= WORD_TO_BYTE(SHR(wValue, 8));
END_IF
m_SetInt:=TRUE;
END_METHOD

//Writes DINT to words nWord, nWord+1 (bytes 2n..2n+3)
METHOD PRIVATE m_SetDint : BOOL
VAR_IN_OUT
	arRaw	: ARRAY[0..127] OF BYTE;
END_VAR
VAR_INPUT
	nWord	: INT;
	nValue	: DINT;
END_VAR
VAR
	dwValue	: DWORD;
	i		: INT;
END_VAR
dwValue:=DINT_TO_DWORD(nValue);
FOR i:=0 TO 3 DO
	IF bSwapBytes THEN;
		arRaw[2*nWord+i]:=DWORD_TO_BYTE(SHR(dwValue, 8*(3-i)));	//most significant byte first
	ELSE;
		arRaw[2*nWord+i]:=DWORD_TO_BYTE(SHR(dwValue, 8*i));		//least significant byte first
	END_IF
END_FOR
m_SetDint:=TRUE;
END_METHOD

END_FUNCTION_BLOCK

// ---- 03 Project/31 AnybusCommunication/FB_Siemens_Sim.TcPOU
//Siemens PLC simulator for tests without the plant. Commissioning tool, off on site.
//Fills the same 128 bytes as the gateway, so FB_Anybus_Interface is tested with its decoding.
//Pumps and hydraulics of the plant are not simulated.
FUNCTION_BLOCK FB_Siemens_Sim
VAR_INPUT
	eMode			: E_Sim_Mode;
	bStart			: BOOL;					//start in eAuto / eQueue
	bStop			: BOOL;					//REQUEST OFF and back to idle
	eFault			: E_Sim_Fault;			//fault to apply
	bFaultOn		: BOOL;					//fault active
	stClient		: ST_Sim_Client := (nClient:=1, eRecipe:=E_Anybus_RecipeType.eFull, eType:=E_Anybus_ClientType.ePipe);
	arQueue			: ARRAY[1..cnQueue] OF ST_Sim_Client;
	stManual		: ST_Anybus_Inputs;		//used in eManual, ALIVE is generated here
	tReplyEmpty		: TIME := T#5S;			//EMPTYING CLIENT -> CLIENT EMPTY
	tReplySprinkler	: TIME := T#3S;			//Sprinkler Request -> Sprinkler State
	tRequestOff		: TIME := T#2S;			//FINISH -> REQUEST OFF
	bSwapBytes		: BOOL := TRUE;			//the same as in FB_Anybus_Interface
END_VAR
VAR_IN_OUT
	arToCip			: ARRAY[0..127] OF BYTE;	//instead of gIO.Anybus_Inputs_Raw
	arFromCip		: ARRAY[0..127] OF BYTE;	//gIO.Anybus_Outputs_Raw
END_VAR
VAR_OUTPUT
	stSend			: ST_Anybus_Inputs;		//sent to CIP, after the fault
	nStep			: INT;					//step of the auto cycle
	nQueuePos		: INT;					//position in arQueue
	bCipReady		: BOOL;					//from CIP
	bCipWorking		: BOOL;
	bCipFinish		: BOOL;
	bCipEmptying	: BOOL;
	bCipPause		: BOOL;
	bCipAlive		: BOOL;
	bCipSprinkler	: BOOL;
	//Text lines of vis_SiemensSim
	sSim			: STRING(120);
	sMode			: STRING(120);
	sClient			: STRING(120);
	sFault			: STRING(120);
	sFromCip		: STRING(120);
	sToCip			: STRING(120);
	sManual			: STRING(120);
	sInterface		: STRING(120);
END_VAR
VAR
	stPlant			: ST_Anybus_Inputs;		//cycle result, before the fault
	bAlive			: BOOL;
	tonAlive		: TON;
	tonEmpty		: TON;
	tonSprinkler	: TON;
	tonOff			: TON;
	tonNext			: TON;
	rtStart			: R_TRIG;
	rtStop			: R_TRIG;
	bSprinklerState	: BOOL;
	nNextShift		: INT;
	i				: INT;
END_VAR
VAR CONSTANT
	cnQueue			: INT := 5;
	cnBadValue		: INT := 99;
	cnIdle			: INT := 0;
	cnWaitReady		: INT := 10;
	cnWaitWorking	: INT := 20;
	cnWaitFinish	: INT := 30;
	cnRequestOff	: INT := 40;
END_VAR

//CIP -> Siemens
bCipReady		:= arFromCip[0].1;
bCipWorking		:= arFromCip[0].2;
bCipFinish		:= arFromCip[0].3;
bCipEmptying	:= arFromCip[0].4;
bCipPause		:= arFromCip[0].6;
bCipAlive		:= arFromCip[0].7;
bCipSprinkler	:= arFromCip[1].0;

//Plant answers
tonEmpty(IN:=bCipEmptying, PT:=tReplyEmpty);
//Sprinkler State follows the request level after tReplySprinkler
tonSprinkler(IN:=bCipSprinkler<>bSprinklerState, PT:=tReplySprinkler);
IF tonSprinkler.Q THEN;
	bSprinklerState:=bCipSprinkler;
END_IF

CASE eMode OF
	E_Sim_Mode.eManual:;
		nStep:=cnIdle;
		stPlant:=stManual;
	E_Sim_Mode.eAuto,
	E_Sim_Mode.eQueue:;
		act_Cycle();
END_CASE
bStart:=FALSE;
bStop:=FALSE;

stSend:=stPlant;
IF eMode<>E_Sim_Mode.eManual THEN;
	stSend.bClientEmpty:=tonEmpty.Q;
	stSend.bSprinklerState:=bSprinklerState;
END_IF
act_Fault();

//ALIVE 0.5 s / 0.5 s
tonAlive(IN:=NOT tonAlive.Q, PT:=T#500MS);
IF tonAlive.Q THEN;
	bAlive:=NOT bAlive;
END_IF
IF NOT (bFaultOn AND eFault=E_Sim_Fault.eAliveStop) THEN;
	stSend.bAlive:=bAlive;
END_IF
act_Status();

//Encode Siemens -> CIP, the layout of FB_Anybus_Interface
IF bFaultOn AND eFault=E_Sim_Fault.eCable THEN;
	FOR i:=0 TO 127 DO
		arToCip[i]:=0;
	END_FOR
	RETURN;
END_IF
arToCip[0].0	:= stSend.bAlarm;
arToCip[0].1	:= stSend.bReady;
arToCip[0].2	:= stSend.bRequestOn;
arToCip[0].3	:= stSend.bRequestOff;
arToCip[0].4	:= stSend.bInletPumpEnable;
arToCip[0].5	:= stSend.bPause;
arToCip[0].6	:= stSend.bClientEmpty;
arToCip[0].7	:= stSend.bAlive;
arToCip[1].0	:= stSend.bSprinklerState;
m_SetInt(arToCip:=arToCip, nWord:=1, nValue:=stSend.nClientId);
m_SetInt(arToCip:=arToCip, nWord:=2, nValue:=stSend.eRecipeType);
m_SetInt(arToCip:=arToCip, nWord:=3, nValue:=stSend.eClientType);
m_SetInt(arToCip:=arToCip, nWord:=4, nValue:=stSend.nNextClient);
m_SetInt(arToCip:=arToCip, nWord:=5, nValue:=stSend.eNextRecipe);
m_SetInt(arToCip:=arToCip, nWord:=6, nValue:=stSend.eNextClientType);

ACTION act_Cycle:
//The plant side of the sequence agreed on 28.10.2026
rtStart(CLK:=bStart);
rtStop(CLK:=bStop);
tonOff(IN:=nStep=cnRequestOff, PT:=tRequestOff);

IF rtStop.Q AND nStep<>cnIdle THEN;
	stPlant.bRequestOn:=FALSE;
	stPlant.bRequestOff:=TRUE;
	nStep:=cnIdle;
END_IF

CASE nStep OF
	cnIdle:;
		stPlant.bReady:=TRUE;
		stPlant.bInletPumpEnable:=TRUE;
		IF rtStart.Q THEN;
			nQueuePos:=1;
			stPlant.bRequestOff:=FALSE;
			m_LoadClient();
			nStep:=cnWaitReady;
		END_IF

	cnWaitReady:;
		IF bCipReady THEN;
			stPlant.bRequestOn:=TRUE;
			stPlant.nClientId:=stPlant.nNextClient;
			stPlant.eRecipeType:=stPlant.eNextRecipe;
			stPlant.eClientType:=stPlant.eNextClientType;
			nStep:=cnWaitWorking;
		END_IF

	cnWaitWorking:;
		IF bCipWorking THEN;
			nStep:=cnWaitFinish;
		END_IF

	cnWaitFinish:;
		IF bCipFinish THEN;
			nStep:=cnRequestOff;
		END_IF

	cnRequestOff:;
		IF tonOff.Q THEN;
			stPlant.bRequestOn:=FALSE;
			stPlant.bRequestOff:=TRUE;
			nQueuePos:=nQueuePos+1;
			IF eMode=E_Sim_Mode.eQueue
			AND nQueuePos<=cnQueue
			AND arQueue[nQueuePos].nClient<>0
			THEN;
				m_LoadClient();
				nStep:=cnWaitReady;
			ELSE;
				nStep:=cnIdle;
			END_IF
		END_IF
END_CASE

//REQUEST OFF is held until CIP drops FINISH
IF stPlant.bRequestOff AND NOT bCipFinish AND NOT bCipWorking THEN;
	stPlant.bRequestOff:=FALSE;
END_IF
END_ACTION

ACTION act_Fault:
tonNext(IN:=bFaultOn AND eFault=E_Sim_Fault.eNextUnstable AND NOT tonNext.Q, PT:=T#1S);
IF tonNext.Q THEN;
	nNextShift:=1-nNextShift;
END_IF
IF NOT bFaultOn THEN;
	nNextShift:=0;
	RETURN;
END_IF

CASE eFault OF
	E_Sim_Fault.ePause:;
		stSend.bPause:=TRUE;
	E_Sim_Fault.eInletOff:;
		stSend.bInletPumpEnable:=FALSE;
	E_Sim_Fault.eRequestDrop:;
		stSend.bRequestOn:=FALSE;
		stSend.bRequestOff:=FALSE;
	E_Sim_Fault.eRequestOff:;
		stSend.bRequestOn:=FALSE;
		stSend.bRequestOff:=TRUE;
	E_Sim_Fault.eConflict:;
		stSend.bRequestOn:=TRUE;
		stSend.bRequestOff:=TRUE;
	E_Sim_Fault.eBadClient:;
		stSend.nClientId:=cnBadValue;
	E_Sim_Fault.eBadRecipe:;
		stSend.eRecipeType:=cnBadValue;
	E_Sim_Fault.eBadType:;
		stSend.eClientType:=cnBadValue;
	E_Sim_Fault.eNextUnstable:;
		stSend.nNextClient:=stSend.nNextClient+nNextShift;
	E_Sim_Fault.eNoClientEmpty:;
		stSend.bClientEmpty:=FALSE;
	E_Sim_Fault.eNoSprinkler:;
		stSend.bSprinklerState:=NOT bCipSprinkler;
	E_Sim_Fault.eReadyOff:;
		stSend.bReady:=FALSE;
END_CASE
END_ACTION

ACTION act_Status:
sSim:=CONCAT('Simulator: ', SEL(g_Anybus.bSimEnable, 'OFF', 'ON'));
sMode:=CONCAT(CONCAT('Mode: ', TO_STRING(eMode)), CONCAT('   step ', TO_STRING(nStep)));
sClient:=CONCAT(CONCAT('Client ', TO_STRING(stClient.nClient)),
	CONCAT(CONCAT('   recipe ', TO_STRING(stClient.eRecipe)), CONCAT('   type ', TO_STRING(stClient.eType))));
sFault:=CONCAT(CONCAT('Fault: ', TO_STRING(eFault)), SEL(bFaultOn, '   armed, not applied', '   APPLIED'));
sFromCip:=CONCAT(CONCAT(CONCAT(CONCAT('CIP: ', m_Bit('READY', bCipReady)), m_Bit('WORKING', bCipWorking)),
	CONCAT(m_Bit('FINISH', bCipFinish), m_Bit('EMPTYING', bCipEmptying))),
	CONCAT(m_Bit('PAUSE', bCipPause), m_Bit('SPRINKLER', bCipSprinkler)));
sToCip:=CONCAT(CONCAT(CONCAT(CONCAT('Plant: ', m_Bit('READY', stSend.bReady)), m_Bit('REQ_ON', stSend.bRequestOn)),
	CONCAT(m_Bit('REQ_OFF', stSend.bRequestOff), m_Bit('INLET', stSend.bInletPumpEnable))),
	CONCAT(CONCAT(m_Bit('PAUSE', stSend.bPause), m_Bit('EMPTY', stSend.bClientEmpty)), m_Bit('SPR_STATE', stSend.bSprinklerState)));
sManual:=CONCAT(CONCAT(CONCAT(CONCAT('Manual: ', m_Bit('READY', stManual.bReady)), m_Bit('REQ_ON', stManual.bRequestOn)),
	CONCAT(m_Bit('REQ_OFF', stManual.bRequestOff), m_Bit('INLET', stManual.bInletPumpEnable))),
	CONCAT(CONCAT(m_Bit('PAUSE', stManual.bPause), m_Bit('EMPTY', stManual.bClientEmpty)), m_Bit('SPR_STATE', stManual.bSprinklerState)));
sInterface:=CONCAT(CONCAT(CONCAT('Interface: ', m_Bit('COMM_OK', g_Anybus.fbAnybus.bCommOk)), CONCAT('request ', TO_STRING(g_Anybus.fbAnybus.eRequest))),
	CONCAT('   alarm ', TO_STRING(g_Anybus.fbAnybus.eAlarm)));
END_ACTION

//Text of one signal for the panel
METHOD PRIVATE m_Bit : STRING(24)
VAR_INPUT
	sName	: STRING(16);
	bValue	: BOOL;
END_VAR
m_Bit:=CONCAT(CONCAT(SEL(bValue, '.', '#'), sName), '  ');
END_METHOD

//NEXT CLIENT for the current position of the cycle
METHOD PRIVATE m_LoadClient : BOOL
VAR
	stNext	: ST_Sim_Client;
END_VAR
IF eMode=E_Sim_Mode.eQueue THEN;
	stNext:=arQueue[nQueuePos];
ELSE;
	stNext:=stClient;
END_IF
stPlant.nNextClient:=stNext.nClient;
stPlant.eNextRecipe:=stNext.eRecipe;
stPlant.eNextClientType:=stNext.eType;
m_LoadClient:=TRUE;
END_METHOD

//Writes INT to word nWord (bytes 2n, 2n+1) of arToCip
METHOD PRIVATE m_SetInt : BOOL
VAR_IN_OUT
	arToCip	: ARRAY[0..127] OF BYTE;
END_VAR
VAR_INPUT
	nWord	: INT;
	nValue	: INT;
END_VAR
VAR
	wValue	: WORD;
END_VAR
wValue:=INT_TO_WORD(nValue);
IF bSwapBytes THEN;
	arToCip[2*nWord]	:= WORD_TO_BYTE(SHR(wValue, 8));
	arToCip[2*nWord+1]	:= WORD_TO_BYTE(wValue);
ELSE;
	arToCip[2*nWord]	:= WORD_TO_BYTE(wValue);
	arToCip[2*nWord+1]	:= WORD_TO_BYTE(SHR(wValue, 8));
END_IF
m_SetInt:=TRUE;
END_METHOD

END_FUNCTION_BLOCK

// ---- 03 Project/31 AnybusCommunication/FB_CIP_Siemens.TcPOU
//Siemens order -> FB_CIP through its existing request buffer, CIP state -> Siemens status.
//Outside the CIP cycle, FB_CIP is not changed. Called in MAIN before act_Call_CIP while g_Anybus.bBridgeEnable.
//One Siemens order at a time: a new one is taken only when the buffer is free (decision B, 02.11.2026).
//Preparing solutions by NEXT (Vadim 02.11.2026, item 8): a local request of FB_CIP, READY = solutions ready.
//Open points are the agent's proposals, see work/vladimir/next_preparation_design.md. Not here yet: flow rate.
//Reaction to ALARM (pause) is temporary, to be confirmed by GAD.
FUNCTION_BLOCK FB_CIP_Siemens
VAR_INPUT
	bWaterOnly		: BOOL;					//commissioning: any order runs as R_Water, no preparation
	bPrepOff		: BOOL := TRUE;			//no preparation by NEXT, READY as soon as CIP is free. TRUE until Vadim decides which chemistry is allowed
	tPrepHold		: TIME := T#30M;		//READY held without circulation, then the preparation is refreshed
	tPrepRetry		: TIME := T#1M;			//new attempt after a preparation that did not reach Done
END_VAR
VAR_OUTPUT
	stStatus		: ST_Anybus_Outputs;	//to g_Anybus.fbAnybus.stStatus
	bActive			: BOOL;					//wash of a Siemens order is in progress
	bFinished		: BOOL;					//wash done, FINISH is held until REQUEST OFF
	bRejected		: BOOL;					//last REQUEST ON was not accepted
	nPrep			: INT;					//preparation state, cnPrep...
	nPrepClient		: INT;					//NEXT CLIENT the solutions are prepared for, 0 = none
	ePrepRecipe		: E_Anybus_RecipeType;	//NEXT RECIPE the solutions are prepared for
END_VAR
VAR
	stReq			: ST_CIP_Request;
	eRecipe			: E_Anybus_RecipeType;
	stBlank			: ST_CIP_Request;
	bTaken			: BOOL;					//our order has reached slot 0 of the buffer
	bStopping		: BOOL;					//cycle reset is running: mRun now would be lost and the order would hang
	tonStopping		: TON;
	bBufferFree		: BOOL;
	bPauseReq		: BOOL;
	bSprinklerReq	: BOOL;
	rtStart			: R_TRIG;				//REQUEST ON while Siemens READY and CIP READY
	tonReadyLost	: TON;					//Siemens READY lost during the wash
	rtPause			: R_TRIG;
	ftPause			: F_TRIG;
	nStage			: INT;
	//Preparation by NEXT
	stPrepReq		: ST_CIP_Request;
	bPrepTaken		: BOOL;					//our local request has reached slot 0 of the buffer
	bPrepMade		: BOOL;					//a local request was needed: refresh after tPrepHold
	nNextNow		: INT;
	eNextNow		: E_Anybus_RecipeType;
	tonPrepHold		: TON;
	tonPrepRetry	: TON;
END_VAR
VAR CONSTANT
	cnNotSupported	: INT := 100;			//order not accepted: CIP busy (proposal)
	cnPrepStart		: INT := 0;				//choose and start the local request when CIP is free
	cnPrepRun		: INT := 1;				//local request in FB_CIP
	cnPrepReady		: INT := 2;				//solutions ready, READY to Siemens
	cnPrepRetry		: INT := 3;				//local request did not reach Done, wait tPrepRetry
	cnPrepWash		: INT := 4;				//Siemens wash, no preparation
END_VAR

bBufferFree:=g_Data.arCIP_RequestBufer[0].eClient=E_CIP_Usage.eNotInUse;
tonStopping(IN:=bStopping, PT:=T#1S);
IF tonStopping.Q THEN;
	bStopping:=FALSE;
END_IF

//Order: only while Siemens READY and CIP READY (solutions prepared). REQUEST ON held from earlier starts the wash
//when both come, a new edge from Siemens is not needed (decisions 02.11.2026). stStatus.bReady of the last cycle
rtStart(CLK:=g_Anybus.fbAnybus.eRequest=E_Anybus_Request.eOn AND g_Anybus.fbAnybus.stIn.bReady AND stStatus.bReady);
IF rtStart.Q
AND NOT bActive
AND NOT bFinished
THEN;
	bRejected:=NOT m_Start();
END_IF

//The way back to Ready clears bRun (_ainit_exit, reset): keep the release until the order leaves Ready
IF (bActive OR nPrep=cnPrepRun)
AND NOT bBufferFree
AND NOT g_Data.b_CIP_Run
AND NOT g_Data.fbCIP.bRun
AND g_Data.fbCIP.eMode<>E_CIP_Mode.eOff
THEN;
	g_Data.fbCIP.mRun();
END_IF

//End of the wash: _aDone_entry frees slot 0
IF bActive THEN;
	IF NOT bBufferFree THEN;
		bTaken:=TRUE;
	ELSIF bTaken THEN;
		bActive:=FALSE;
		bTaken:=FALSE;
		bFinished:=TRUE;
	END_IF
END_IF

//REQUEST OFF: confirms FINISH or stops the wash
IF g_Anybus.fbAnybus.eRequest=E_Anybus_Request.eOff
OR g_Anybus.fbAnybus.eRequest=E_Anybus_Request.eConflict
THEN;
	bFinished:=FALSE;
	bRejected:=FALSE;
	IF bActive THEN;
		m_Stop();
	END_IF
END_IF

//Preparation by NEXT: free CIP prepares the solutions for the accepted NEXT, READY when done, refresh after tPrepHold.
//A change of NEXT stops the preparation and starts it for the new NEXT
IF g_Anybus.fbAnybus.bNextValid THEN;
	nNextNow:=g_Anybus.fbAnybus.nNextClient;
	eNextNow:=g_Anybus.fbAnybus.eNextRecipe;
ELSE;
	nNextNow:=0;
	eNextNow:=E_Anybus_RecipeType.eNone;
END_IF
IF bActive OR bFinished THEN;
	nPrep:=cnPrepWash;
ELSIF (nPrep=cnPrepRun OR nPrep=cnPrepReady OR nPrep=cnPrepRetry)
AND (nNextNow<>nPrepClient OR eNextNow<>ePrepRecipe)
THEN;
	IF nPrep=cnPrepRun THEN;
		m_PrepStop();
	END_IF
	nPrep:=cnPrepStart;
END_IF
tonPrepHold(IN:=nPrep=cnPrepReady AND bPrepMade, PT:=tPrepHold);
tonPrepRetry(IN:=nPrep=cnPrepRetry, PT:=tPrepRetry);
CASE nPrep OF
	cnPrepWash:;
		IF NOT bActive AND NOT bFinished THEN;
			nPrep:=cnPrepStart;
		END_IF

	cnPrepStart:;
		IF bBufferFree
		AND NOT bStopping
		AND NOT g_Data.fbCIP.bRun
		AND g_Data.fbCIP.SFCCurrentStep='Ready'
		AND g_Data.fbCIP.eMode<>E_CIP_Mode.eOff
		THEN;
			nPrepClient:=nNextNow;
			ePrepRecipe:=eNextNow;
			bPrepMade:=NOT bPrepOff AND NOT bWaterOnly AND m_PrepRequest();
			IF bPrepMade THEN;
				g_Data.fbCIP.m_TakePosInCIPBuffer(stCIP_Request:=stPrepReq);
				g_Data.fbCIP.mRun();
				bPrepTaken:=FALSE;
				nPrep:=cnPrepRun;
			ELSE;
				nPrep:=cnPrepReady;
			END_IF
		END_IF

	cnPrepRun:;
		//_aDone_entry frees slot 0; freed without Done = stopped from outside
		IF NOT bBufferFree THEN;
			bPrepTaken:=TRUE;
		ELSIF bPrepTaken THEN;
			bPrepTaken:=FALSE;
			IF g_Data.fbCIP.bDone THEN;
				nPrep:=cnPrepReady;
			ELSE;
				nPrep:=cnPrepRetry;
			END_IF
		END_IF

	cnPrepReady:;
		IF tonPrepHold.Q THEN;
			nPrep:=cnPrepStart;
		END_IF

	cnPrepRetry:;
		IF tonPrepRetry.Q THEN;
			nPrep:=cnPrepStart;
		END_IF
END_CASE

//Recipe of the local preparation in FB_CIP: the client of the wash, the NEXT client while preparing, else Local
IF bActive THEN;
	g_Data.fbCIP.nLocalRecipe:=stReq.nClientId;
ELSIF nPrep=cnPrepRun THEN;
	g_Data.fbCIP.nLocalRecipe:=nPrepClient;
ELSE;
	g_Data.fbCIP.nLocalRecipe:=0;
END_IF

//Pause, the existing CIP zone Pause / Play. Play comes by itself when all causes are gone (decision 02.11.2026)
tonReadyLost(IN:=bActive AND NOT g_Anybus.fbAnybus.stIn.bReady, PT:=T#1S);
bPauseReq:=bActive AND (
	g_Anybus.fbAnybus.eRequest=E_Anybus_Request.eNone
	OR tonReadyLost.Q
	OR g_Anybus.fbAnybus.stIn.bPause
	OR g_Anybus.fbAnybus.stIn.bAlarm
	OR NOT g_Anybus.fbAnybus.stIn.bInletPumpEnable);
rtPause(CLK:=bPauseReq);
ftPause(CLK:=bPauseReq);
IF rtPause.Q THEN;
	stOper[E_ModeZone.eCIP].bSetPause:=TRUE;
END_IF
IF ftPause.Q THEN;
	stOper[E_ModeZone.eCIP].bSetPlay:=TRUE;
END_IF

//Status
stStatus.bReady:=TRUE
	AND NOT bActive
	AND NOT bFinished
	AND NOT bStopping
	AND bBufferFree
	AND NOT g_Data.fbCIP.bRun
	AND g_Data.fbCIP.SFCCurrentStep='Ready'
	AND g_Data.fbCIP.eMode<>E_CIP_Mode.eOff
	AND g_Anybus.fbAnybus.bCommOk
	AND nPrep=cnPrepReady;
stStatus.bWorking:=bActive;
//SENDING PUMP WORKING: the CIP sending pump P1001 runs during the Siemens wash, for indication in the plant
stStatus.bSendingPump:=bActive AND g_Pump.fbPump[E_Pump_List.P1001].bRun;
//EMPTYING CLIENT: Tank on a Tank_LowLevel step, the steps wait for CLIENT EMPTY
stStatus.bEmptyingClient:=bActive
	AND stReq.eClientType=E_Anybus_ClientType.eTank
	AND FIND(g_Data.fbCIP.SFCCurrentStep, 'Tank_LowLevel')>0;
//Sprinkler: on from CIPx_Conn_Sprinkler until FB_CIP leaves the spray ball, off until Siemens confirms.
//bSprinkler alone is too early: the mix-proof steps set it before CIP2 and CIP4
IF NOT bActive OR NOT g_Data.fbCIP.bSprinkler THEN;
	bSprinklerReq:=FALSE;
END_IF
IF bActive AND FIND(g_Data.fbCIP.SFCCurrentStep, 'Conn_Sprinkler')>0 THEN;
	bSprinklerReq:=TRUE;
END_IF
//One level bit: 0 asks Siemens back to the pipe, Sprinkler State 0 confirms (Vadim 02.11.2026, items 7-8)
stStatus.bSprinklerRequest:=bSprinklerReq;
stStatus.bFinish:=bFinished;
stStatus.bPause:=bActive AND stOper[E_ModeZone.eCIP].iActOperation=E_OperationButtons.ePauseAll;
stStatus.eActualMedia:=m_Media();
//Progress of the current medium in seconds (proposal, to be confirmed by Vadim): circulation timer of FB_CIP,
//reset at the start of each medium. Remaining time to the next stage = recipe - actual
IF bActive THEN;
	stStatus.nRecipeProgress:=TIME_TO_DINT(g_Data.fbCIP.tonr_CIP_Condition.PT)/1000;
	stStatus.nActualProgress:=TIME_TO_DINT(g_Data.fbCIP.tonr_CIP_Condition.ET)/1000;
ELSE;
	stStatus.nRecipeProgress:=0;
	stStatus.nActualProgress:=0;
END_IF
IF bActive OR bFinished THEN;
	stStatus.nActiveClient:=stReq.nClientId;
	stStatus.eActiveRecipe:=eRecipe;
ELSE;
	stStatus.nActiveClient:=0;
	stStatus.eActiveRecipe:=E_Anybus_RecipeType.eNone;
END_IF
IF bRejected THEN;
	stStatus.nAlarmCode:=cnNotSupported;
ELSE;
	stStatus.nAlarmCode:=0;
END_IF

//TRUE: the order is in the CIP buffer and the cycle is released
METHOD PRIVATE m_Start : BOOL
//Not before Ready: after a stop the way back to Ready (valves, client drain) takes more than bStopping,
//_aReady_exit would be missed and eCIP_State of the order not taken
IF NOT g_Anybus.fbAnybus.bCurrentValid
OR bStopping
OR NOT bBufferFree
OR g_Data.fbCIP.bRun
OR g_Data.fbCIP.SFCCurrentStep<>'Ready'
OR g_Data.fbCIP.eMode=E_CIP_Mode.eOff
THEN;
	RETURN;
END_IF

//GAD wash type -> CIP type and first stage, table of 02.11.2026
CASE g_Anybus.fbAnybus.stIn.eRecipeType OF
	E_Anybus_RecipeType.eFlushOnly:;
		stReq.eType:=E_CIP_Type.R_Water;
		stReq.eStartState:=E_Element_State_Long.eNotClean;
	E_Anybus_RecipeType.eDetergent:;
		stReq.eType:=E_CIP_Type.Detergent;
		stReq.eStartState:=E_Element_State_Long.eNotClean;
	E_Anybus_RecipeType.eDetergentOnly:;
		stReq.eType:=E_CIP_Type.Detergent;
		stReq.eStartState:=E_Element_State_Long.eCIP_1_Rinzed;
	E_Anybus_RecipeType.eDisinfectionOnly:;
		stReq.eType:=E_CIP_Type.Full;
		stReq.eStartState:=E_Element_State_Long.eCIP_3_Deterged_Clean;
	E_Anybus_RecipeType.eDetergentDisinfection:;
		stReq.eType:=E_CIP_Type.Full;
		stReq.eStartState:=E_Element_State_Long.eCIP_1_Rinzed;
	E_Anybus_RecipeType.eFull:;
		stReq.eType:=E_CIP_Type.Full;
		stReq.eStartState:=E_Element_State_Long.eNotClean;
ELSE;
	RETURN;
END_CASE
IF bWaterOnly THEN;
	stReq.eType:=E_CIP_Type.R_Water;
	stReq.eStartState:=E_Element_State_Long.eNotClean;
END_IF
eRecipe:=g_Anybus.fbAnybus.stIn.eRecipeType;
stReq.eClient:=E_CIP_Usage.eExternal;
stReq.nClientId:=g_Anybus.fbAnybus.stIn.nClientId;
stReq.eClientType:=g_Anybus.fbAnybus.stIn.eClientType;

g_Data.fbCIP.m_TakePosInCIPBuffer(stCIP_Request:=stReq);
g_Data.fbCIP.mRun();
bActive:=TRUE;
bTaken:=FALSE;
m_Start:=TRUE;
END_METHOD

//REQUEST OFF during the wash. Not bStopResetAll: it puts the CIP zone to Manual and Pause, the next order would not run
METHOD PRIVATE m_Stop : BOOL
g_Data.arCIP_RequestBufer[0]:=stBlank;
g_Data.fbCIP.mResetCycle();
bStopping:=TRUE;
bActive:=FALSE;
bTaken:=FALSE;
m_Stop:=TRUE;
END_METHOD

//Local request for ePrepRecipe, table of Vadim 02.11.2026. FALSE: no solution is needed (no NEXT, Flush_Only).
//The start state is set as in the table, FB_CIP takes it for local requests only with item 7 (later)
METHOD PRIVATE m_PrepRequest : BOOL
stPrepReq:=stBlank;
stPrepReq.eClient:=E_CIP_Usage.eLocal;
CASE ePrepRecipe OF
	E_Anybus_RecipeType.eDetergent, E_Anybus_RecipeType.eDetergentOnly:;
		//T92
		stPrepReq.eType:=E_CIP_Type.Detergent;
		stPrepReq.eStartState:=E_Element_State_Long.eCIP_1_Rinzed;
	E_Anybus_RecipeType.eDisinfectionOnly:;
		//T91
		stPrepReq.eType:=E_CIP_Type.Full;
		stPrepReq.eStartState:=E_Element_State_Long.eCIP_3_Deterged_Clean;
	E_Anybus_RecipeType.eDetergentDisinfection, E_Anybus_RecipeType.eFull:;
		//T92 and T91
		stPrepReq.eType:=E_CIP_Type.Full;
		stPrepReq.eStartState:=E_Element_State_Long.eCIP_1_Rinzed;
ELSE;
	RETURN;
END_CASE
m_PrepRequest:=TRUE;
END_METHOD

//NEXT changed during the preparation: the same stop as on REQUEST OFF
METHOD PRIVATE m_PrepStop : BOOL
g_Data.arCIP_RequestBufer[0]:=stBlank;
g_Data.fbCIP.mResetCycle();
bStopping:=TRUE;
bPrepTaken:=FALSE;
m_PrepStop:=TRUE;
END_METHOD

//Actual Media by the dashboard stage of FB_CIP
METHOD PRIVATE m_Media : E_Anybus_Media
m_Media:=E_Anybus_Media.eNone;
IF NOT bActive THEN;
	RETURN;
END_IF
nStage:=TO_INT(g_HMI.eCIP_DashStage_actual);
CASE nStage OF
	1..2:;
		m_Media:=E_Anybus_Media.eFirstWater;
	3..7:;
		m_Media:=E_Anybus_Media.eSoda;
	8..11:;
		m_Media:=E_Anybus_Media.eIntermediateWater;
	12..16:;
		m_Media:=E_Anybus_Media.eDisinfection;
	17..20:;
		m_Media:=E_Anybus_Media.eLastWater;
END_CASE
END_METHOD

END_FUNCTION_BLOCK

// ---- 00 Library/00-General/CheckBounds.TcPOU
FUNCTION CheckBounds : DINT
VAR_INPUT
	index, lower, upper : DINT;
END_VAR
VAR
END_VAR

IF index<lower THEN
	CheckBounds := lower;
	Errors:=Errors+1;
ELSIF index>upper THEN
	CheckBounds := upper;
	Errors:=Errors+1;
ELSE
	CheckBounds := index;
END_IF

END_FUNCTION

// ---- 00 Library/00-General/TimeAndDate/FUN_DeltaTime.TcPOU
FUNCTION FUN_DeltaTime : STRING
VAR_INPUT
    //stSystemTime : TimeStruct;
    stStartTime  : TimeStruct;	
END_VAR
VAR
    dtSystemTime : DT;
    dtStartTime  : DT;
    deltaTime    : TIME;
    hours        : INT;
    minutes      : INT;
    milliseconds : INT;
    sDeltaTime   : STRING;	
END_VAR

// Convert TimeStruct to DT
dtSystemTime := SYSTEMTIME_TO_DT(stSystemTime);
dtStartTime  := SYSTEMTIME_TO_DT(stStartTime);

// Calculate the delta time
deltaTime := TO_TIME(dtSystemTime - dtStartTime);

// Extract hours, minutes, and milliseconds
hours := INT_TO_DINT(deltaTime / T#1H);
minutes := INT_TO_DINT((deltaTime MOD T#1H) / T#1M);
milliseconds := INT_TO_DINT((deltaTime MOD T#1M) / T#1MS);

// Format the string
sDeltaTime := CONCAT(CONCAT(CONCAT(CONCAT(INT_TO_STRING(hours), ':'), INT_TO_STRING(minutes)), ':'), INT_TO_STRING(milliseconds));

FUN_DeltaTime := sDeltaTime;

END_FUNCTION

// ---- 00 Library/04 Recipe/OLD/prg_RecipeManager.TcPOU
PROGRAM prg_RecipeManager
VAR
	fbRecipe: RecipeManCommands;
	LastError: DWORD;
	LastInfo: InfoValues;

	bCheckError: BOOL;
	bResetError: BOOL;
	bInit: BOOL;
END_VAR


IF bCheckError THEN;
	//bCheckError:=FALSE;
	LastError:=fbRecipe.GetLastError();
	LastInfo:=fbRecipe.GetLastInfo();
END_IF

IF bResetError THEN;
	bResetError:=FALSE;
	LastError:=fbRecipe.ResetLastError();
	LastError:=fbRecipe.ReloadRecipes(RecipeDefinitionName:='');
	
END_IF

IF bInit THEN;
	bInit:=FALSE;
	LastError:=fbRecipe.ResetLastInfo();
END_IF

END_PROGRAM

// ---- 00 Library/04-Messages/FB_PrintErrMessageByID_ST_Cycle.TcPOU
FUNCTION_BLOCK FB_PrintErrMessageByID_ST_Cycle
VAR_INPUT
	pstCycle			:POINTER TO ST_BasicCycle;
	sActErrorID			: STRING;
	ErrorToPrint		: STRING;
	iFB_Num				: INT:=0;
	sFB_ModuleDescription	:STRING(30):='';
	bResumeAll		: BOOL;
END_VAR
VAR_OUTPUT
END_VAR
VAR
	cFound				: INT;
	i					: INT;
	iFound				: INT;
	//r_trigPrintMessage	: R_TRIG;
	bNewMeasege			: BOOL;
	sActErrorID_AA		: STRING;
	iErrorID_Flag		: INT;
	sAA					: STRING;
	sActErrorID_Message	: STRING;
	iAAPos				: INT;
	rtrig1				: R_TRIG;
	
	sLastErrorID: STRING;
	j: INT;
END_VAR


IF pstCycle^.bFault THEN
	IF sActErrorID<>'000x000x000'  AND sActErrorID<>'' THEN //to print or not to print the massage???
		sLastErrorID:=sActErrorID;
		bNewMeasege:=TRUE;
		FOR i:=1 TO 100 DO
			IF Buffer_Act_Message[i].sErrID=sActErrorID THEN;
				IF Buffer_Act_Message[i].sModuleDescription = sFB_ModuleDescription THEN
					bNewMeasege:=FALSE;
					EXIT;
				END_IF
			END_IF
		END_FOR
	ELSE
		bNewMeasege:=FALSE;
	END_IF
	
	IF bNewMeasege AND NOT bResumeAll THEN;
		FOR i:=100 TO 2 BY -1 DO
			Buffer_Act_Message[i].sDateTime:=Buffer_Act_Message[i-1].sDateTime;
			Buffer_Act_Message[i].sErrID:=Buffer_Act_Message[i-1].sErrID;
			Buffer_Act_Message[i].sErrorMessage:=Buffer_Act_Message[i-1].sErrorMessage;
			Buffer_Act_Message[i].sLevel:=Buffer_Act_Message[i-1].sLevel;
			Buffer_Act_Message[i].sModuleDescription:=Buffer_Act_Message[i-1].sModuleDescription;
		END_FOR
		
		Buffer_Act_Message[1].sDateTime:=prg_RealClock.sRealTime_Date;
		Buffer_Act_Message[1].sErrID:=sActErrorID;
		Buffer_Act_Message[1].sModuleDescription:=sFB_ModuleDescription;

		IF sActErrorID='000x000x999' THEN;
			Buffer_Act_Message[1].sErrorMessage:=CONCAT('Cycle message: ',ErrorToPrint);
		ELSE
			cFound:=0;
			FOR i:=1 TO C_Max_ErrorList DO
				IF ar_ErrorList[i,eErrID]=sActErrorID THEN
					iFound:=i;
					ar_ErrorActive[iFound]:=TRUE;
					cFound:=cFound+1;
				END_IF
			END_FOR
	
			IF cFound=1 THEN;
				Buffer_Act_Message[1].sErrorMessage:=ar_ErrorList[iFound,eErrMeassage];	(*	Error from the List	*)
				pstCycle^.sFailedMessage := Buffer_Act_Message[1].sErrorMessage;
				Buffer_Act_Message[1].sLevel:=ar_ErrorList[iFound,eErrLevel];	(*	Error Level from the List	*)
			ELSIF cFound=0 THEN; //(*	Error ID not Foud on the List	*)
				//Buffer_Act_Message[1].sErrorMessage:='Error ID not found on the "Error List"';
				Buffer_Act_Message[1].sErrorMessage:=CONCAT('Cycle message[1]: ',ErrorToPrint);
				Buffer_Act_Message[1].sLevel:='Error';
			ELSIF cFound>1 THEN; //(*	More then one Errors Foud with the same  ID		*)
				//Buffer_Act_Message[1].sErrorMessage:='More then one error with the same ID  found on the "Error list"';
				Buffer_Act_Message[1].sErrorMessage:=CONCAT('Cycle message[2]: ',ErrorToPrint);
				Buffer_Act_Message[1].sLevel:='Error';
			END_IF
		END_IF
		FUN_Write_Line_To_History();
	END_IF
	
	
	IF bResumeAll THEN
		sActErrorID:='';
	END_IF
	
END_IF

(*
//for delete message if no fault
rtrig1(CLK:= NOT pstCycle^.bFault, Q=> );
IF rtrig1.Q THEN  // if cycle not in pause
	FOR i:= 2 TO 100 DO //loop for search 
		IF Buffer_Act_Message[i-1].sErrID = sLastErrorID THEN // search if last error id = buffer which it error table.
			FOR j:= i TO 100 DO //if found message id then delete it.
				Buffer_Act_Message[j-1]:=Buffer_Act_Message[j];//delete
			END_FOR
		END_IF
	END_FOR
END_IF
*)

END_FUNCTION_BLOCK

// ---- 00 Library/07 Errors/FB_Error_Handle.TcPOU
FUNCTION_BLOCK FB_Error_Handle
VAR_INPUT
	bError: BOOL;
	sErrID: STRING;
END_VAR
VAR_OUTPUT
END_VAR
VAR
	fbFormat: FB_FormatString;
END_VAR
VAR_IN_OUT
	error_code: STRING;

END_VAR



IF bError 
AND error_code=''
THEN;
	error_code:=sErrID;
END_IF

IF NOT bError 
AND error_code=sErrID
THEN;
	error_code:='';
END_IF

METHOD m_GetAxisErr : STRING(4)
VAR_INPUT
	stDevErr_H				: ST_DeviceErrorHandeling;
END_VAR
VAR_OUTPUT
	sMessage: STRING;
END_VAR

VAR
	ErrID_xx: STRING(2);
END_VAR
IF bError 
AND error_code=''
THEN;
	fbFormat(sFormat:='%0.2d' ,arg1:=F_INT(stDevErr_H.iObjectID),sOut=>ErrID_xx);
	m_GetAxisErr:=CONCAT('23',ErrID_xx);
	sMessage:=stDevErr_H.sObjectName;
ELSE;
	m_GetAxisErr:='';
END_IF
END_METHOD

METHOD m_GetPistonErr : STRING(4)
VAR_INPUT
	stDevErr_H				: ST_DeviceErrorHandeling;
END_VAR
VAR_OUTPUT
	sMessage: STRING;
END_VAR

VAR
	ErrID_xx: STRING(2);
END_VAR
IF bError 
AND error_code=''
THEN;
	fbFormat(sFormat:='%0.2d' ,arg1:=F_INT(stDevErr_H.iObjectID),sOut=>ErrID_xx);
	m_GetPistonErr:=CONCAT('22',ErrID_xx);
	sMessage:=stDevErr_H.sObjectName;
ELSE;
	m_GetPistonErr:='';
END_IF
END_METHOD

END_FUNCTION_BLOCK

// ---- 00 Library/10 Utils/DutyCycle/FB_DutyCycle.TcPOU
FUNCTION_BLOCK FB_DutyCycle
VAR_INPUT
	bEnable		: BOOL;
	fBaseTime	: REAL:=5.0; // [sec] min>0
	fOn_Duty	: REAL:=10.0; //min =0, max=100
END_VAR
VAR_OUTPUT
	bOut: BOOL;
END_VAR
VAR
	tBaseTime: TIME;
	ton_OnDuty: TON;
	fOnTime: REAL;
	tOnTime: TIME;
END_VAR


tBaseTime:=REAL_TO_TIME(fBaseTime*1000);
ton_OnDuty(PT:=tBaseTime,IN:=NOT ton_OnDuty.Q AND bEnable);

IF fOn_Duty<0 THEN;
	fOn_Duty:=0;
ELSIF fOn_Duty>100 THEN;
	fOn_Duty:=1000;
END_IF
	
fOnTime:=fBaseTime*fOn_Duty/100.0;
tOnTime:=REAL_TO_TIME(fOnTime*1000);

IF bEnable THEN;
	IF fOn_Duty<=0 THEN;
		bOut:=FALSE;
	ELSIF fOn_Duty>=100 THEN;
		bOut:=TRUE;
	ELSE;
		IF ton_OnDuty.ET<tOnTime THEN;
			bOut:=TRUE;
		ELSE
			bOut:=FALSE;
		END_IF		
	END_IF	
ELSE;
	bOut:=FALSE;
END_IF

END_FUNCTION_BLOCK

// ---- 00 Library/10 Utils/fun_LrealToString.TcPOU
FUNCTION fun_LrealToString : STRING
VAR_INPUT
	iDigits	: INT:=2;
	fVar	: LREAL;
END_VAR
VAR
	iDigitsLocal: INT;

	fTemp: LREAL;
	fMult: LREAL;
	
	fbFormat: FB_FormatString;	

END_VAR

IF iDigits<0 THEN;
	iDigitsLocal:=0;
ELSIF iDigits>6 THEN;
	iDigitsLocal:=6; 
ELSE
	iDigitsLocal:=iDigits;	
END_IF

// this vertion solve the case then the result is 2.0-e2 instade of 0.02
CASE iDigitsLocal OF
	0:;fbFormat(sFormat:='%.0f' ,arg1:=F_LREAL(fVar),sOut=>fun_LrealToString);
	1:;fbFormat(sFormat:='%.1f' ,arg1:=F_LREAL(fVar),sOut=>fun_LrealToString);
	2:;fbFormat(sFormat:='%.2f' ,arg1:=F_LREAL(fVar),sOut=>fun_LrealToString);
	3:;fbFormat(sFormat:='%.3f' ,arg1:=F_LREAL(fVar),sOut=>fun_LrealToString);
	4:;fbFormat(sFormat:='%.4f' ,arg1:=F_LREAL(fVar),sOut=>fun_LrealToString);
	5:;fbFormat(sFormat:='%.5f' ,arg1:=F_LREAL(fVar),sOut=>fun_LrealToString);
	6:;fbFormat(sFormat:='%.6f' ,arg1:=F_LREAL(fVar),sOut=>fun_LrealToString);
END_CASE

(* OLD Version
CASE iDigitsLocal OF
	0:;fMult:=1;
	1:;fMult:=10;
	2:;fMult:=100;
	3:;fMult:=1000;
	4:;fMult:=10000;
	5:;fMult:=100000;
	6:;fMult:=1000000;
END_CASE

fTemp:=TRUNC(fVar*fMult);
IF iDigitsLocal=0 THEN;
	fun_LrealToString:=DINT_TO_STRING(TRUNC(fVar));
ELSE;
	fun_LrealToString:=LREAL_TO_STRING(fTemp/fMult);	
END_IF
*)

END_FUNCTION

// ---- 00 Library/10 Utils/F_TimeRatio.TcPOU
FUNCTION F_TimeRatio : INT
VAR_INPUT
	t1: TIME;
	t2: TIME;

END_VAR
VAR
	udi_t1: UDINT;
	udi_t2: UDINT;

	ratio: REAL;
END_VAR


udi_t1:=TIME_TO_UDINT(t1);
udi_t2:=TIME_TO_UDINT(t2);

IF udi_t2>0 THEN;
	ratio:=udi_t1/udi_t2;
END_IF

END_FUNCTION

// ---- 01 Instance/04-Messages/Prg_Filter_Messages.TcPOU
PROGRAM Prg_Filter_Messages
VAR
	sSearchMessage		: STRING;
	i					: INT;
	d					: INT;
	stFilter			: stMessageFormat;
	stLastFilter		: stMessageFormat;
	T1					: TON;
	bFilter				: BOOL;
END_VAR


IF stFilter.sErrID<>stLastFilter.sErrID
OR  stFilter.sLevel <>stLastFilter.sLevel
OR  stFilter.sModuleDescription <>stLastFilter.sModuleDescription
OR  stFilter.sErrorMessage<>stLastFilter.sErrorMessage THEN

	FOR i:=1000 TO 1 BY -1 DO
		Buffer_Search_Messages[i].sDateTime:='';
		Buffer_Search_Messages[i].sErrID:='';
		Buffer_Search_Messages[i].sErrorMessage:='';
		Buffer_Search_Messages[i].sLevel:='';
		Buffer_Search_Messages[i].sModuleDescription:='';
	END_FOR
	bFilter:=TRUE;
ELSE
	bFilter:=FALSE;
END_IF




T1(IN:=bFilter , PT:=T#300MS , Q=> , ET=> );
IF T1.Q THEN
	d:=2;
	FOR i:=1 TO 1000 DO
			IF (Buffer_Act_History[i].sErrID=stFilter.sErrID OR stFilter.sErrID='')
			AND (Buffer_Act_History[i].sLevel=stFilter.sLevel OR stFilter.sLevel='')
			AND (Buffer_Act_History[i].sErrorMessage=stFilter.sErrorMessage OR stFilter.sErrorMessage='')
			AND (Buffer_Act_History[i].sModuleDescription=stFilter.sModuleDescription OR stFilter.sModuleDescription='')THEN
				Buffer_Search_Messages[d]:=Buffer_Act_History[i];
				d:=d+1;
			END_IF
	END_FOR
	
	
ELSE

FOR i:=1000 TO 2 BY -1 DO
	Buffer_Search_Messages[i]:=Buffer_Act_History[i-1];
END_FOR

END_IF

END_PROGRAM

// ---- 01 Instance/07-Mode/prg_HMI_OperationLock.TcPOU
PROGRAM prg_HMI_OperationLock
VAR
	b_LockIndex: BOOL;
	b_LockLoad: BOOL;
	b_LockUnload: BOOL;
	b_LockManip: BOOL;
END_VAR

IF stModeMain.iActMode= 2 AND prg_User.actUser< 3 THEN
   b_LockIndex := TRUE;
ELSE
   b_LockIndex := FALSE;
END_IF

END_PROGRAM

// ---- 00 Library/01 Piston/TextList_Piston_Recipe_State.TcTLO
TEXTLIST TextList_Piston_Recipe_State
  0 = ' '
  1 = 'Open'
  2 = 'Close'
   = ''
END_TEXTLIST

// ---- 00 Library/01 Piston/TextList_Piston_Recipe_State_CloseOpen.TcTLO
TEXTLIST TextList_Piston_Recipe_State_CloseOpen
  0 = ' '
  1 = 'Close'
  2 = 'Open'
   = ''
END_TEXTLIST

// ---- 00 Library/01 Piston/TextList_Piston_Recipe_State_DownUp.TcTLO
TEXTLIST TextList_Piston_Recipe_State_DownUp
  0 = ' '
  1 = 'Down'
  2 = 'Up'
   = ''
END_TEXTLIST

// ---- 00 Library/01 Piston/TextList_Piston_Recipe_State_InOut.TcTLO
TEXTLIST TextList_Piston_Recipe_State_InOut
  0 = ' '
  1 = 'In'
  2 = 'Out'
   = ''
END_TEXTLIST

// ---- 00 Library/01 Piston/TextList_Piston_Recipe_State_OnOff.TcTLO
TEXTLIST TextList_Piston_Recipe_State_OnOff
  0 = ' '
  1 = 'On'
  2 = 'Off'
   = ''
END_TEXTLIST

// ---- 00 Library/01 Piston/TextList_Piston_Recipe_State_OpenClose.TcTLO
TEXTLIST TextList_Piston_Recipe_State_OpenClose
  0 = ' '
  1 = 'Open'
  2 = 'Close'
   = ''
END_TEXTLIST

// ---- 00 Library/01 Piston/TextList_Piston_Recipe_State_UpDown.TcTLO
TEXTLIST TextList_Piston_Recipe_State_UpDown
  0 = ' '
  1 = 'Up'
  2 = 'Down'
   = ''
END_TEXTLIST

// ---- 00 Library/01 Piston/VISU/vis_Piston_Control1.TcVIS
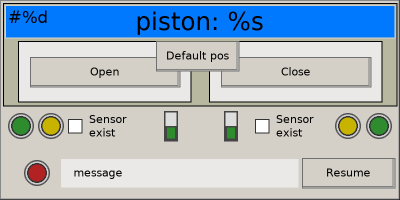
VISUALIZATION vis_Piston_Control1  // 400x200
VAR_IN_OUT
	stPis: ST_Piston;
END_VAR
    Rectangle (0,0 400x200)
    Rectangle (3,3 394x103), colour toggle: NOT stPis.b_Enable
    Rectangle (18,41 173x61), colour toggle: stPis.st_Open
    Rectangle (209,41 173x61), colour toggle: stPis.st_Close
    Button (30,57 150x30), "Open", colour toggle: stPis.req_Open, input disabled if: stPis.b_DeactivateMan OR NOT stPis.b_InterLock_Open
        toggle stPis.req_OpenMan
    Button (221,57 150x30), "Close", colour toggle: stPis.req_Close, input disabled if: stPis.b_DeactivateMan OR NOT stPis.b_InterLock_Close
        toggle stPis.req_CloseMan
    DipSwitch (156,111 30x30), tooltip "Open Sensor state", variable: stPis.sen_Open, invisible if: NOT stPis.sen_Open_Exist, behaviour: TOGGLE, style: Switch-DipSwitch-Green
    DipSwitch (216,111 30x30), tooltip "Close Sensor state", variable: stPis.sen_Close, invisible if: NOT stPis.sen_Close_Exist, behaviour: TOGGLE, style: Switch-DipSwitch-Green
    Checkbox (66,108 99x36), "Sensor exist", variable: stPis.sen_Open_Exist
    Checkbox (253,108 99x36), "Sensor exist", variable: stPis.sen_Close_Exist
    Lamp1 (6,111 30x30), tooltip "Open sensor", variable: stPis.sen_Open, invisible if: NOT stPis.sen_Open_Exist, style: Lamp-Lamp1-Green
    Lamp1 (333,111 30x30), tooltip "Close valve", variable: stPis.valve_Close, style: Lamp-Lamp1-Yellow
    Lamp1 (22,158 30x30), tooltip "Error", variable: stPis.b_Error, style: Lamp-Lamp1-Red
    Textfield (60,158 239x30), "message"
    Button (302,158 93x30), "Resume", colour toggle: stPis.b_Error
        toggle stPis.b_Resume
    Button (156,41 83x30), "Default pos", colour toggle: stPis.req_DefaultPos, input disabled if: stPis.b_DeactivateMan
        toggle stPis.req_DefaultPos
    Textfield (5,5 390x33), "piston: %s", text variable: stPis.sName
    Textfield (5,7 42x21), "#%d", text variable: stPis.iPisNum
    Lamp1 (36,111 30x30), tooltip "Open valve", variable: stPis.valve_Open, style: Lamp-Lamp1-Yellow
    Lamp1 (364,111 30x30), tooltip "Close sensor", variable: stPis.sen_Close, invisible if: NOT stPis.sen_Close_Exist, style: Lamp-Lamp1-Green
END_VISUALIZATION

// ---- 00 Library/01 Piston/VISU/vis_Piston_Control1_Compact.TcVIS
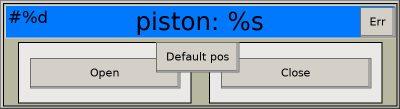
VISUALIZATION vis_Piston_Control1_Compact  // 400x109
VAR_IN_OUT
	stPis: ST_Piston;
END_VAR
    Rectangle (0,0 400x109)
    Rectangle (3,3 394x103), colour toggle: NOT stPis.b_Enable
    Rectangle (18,42 173x61), colour toggle: stPis.st_Open
    Rectangle (209,42 173x61), colour toggle: stPis.st_Close
    Button (30,58 150x30), "Open", colour toggle: stPis.req_Open, input disabled if: stPis.b_DeactivateMan OR NOT stPis.b_InterLock_Open
        toggle stPis.req_OpenMan
    Button (221,58 150x30), "Close", colour toggle: stPis.req_Close, input disabled if: stPis.b_DeactivateMan OR NOT stPis.b_InterLock_Close
        toggle stPis.req_CloseMan
    Button (156,42 83x30), "Default pos", colour toggle: stPis.req_DefaultPos, input disabled if: stPis.b_DeactivateMan
        toggle stPis.req_DefaultPos
    Textfield (5,5 390x33), "piston: %s", text variable: stPis.sName
    Textfield (5,7 42x21), "#%d", text variable: stPis.iPisNum
    Button (360,7 35x30), "Err", colour toggle: stPis.b_Error
        toggle stPis.b_Resume
END_VISUALIZATION

// ---- 00 Library/01 Piston/VISU/vis_Piston_Control2_CloseOpen.TcVIS
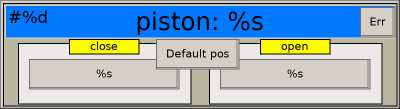
VISUALIZATION vis_Piston_Control2_CloseOpen  // 400x109
VAR_IN_OUT
	stPis			: ST_Piston;
END_VAR
VAR_INPUT
	sLable_Open		: STRING:='lable open';
	sLable_Close	: STRING:='lable close';
END_VAR
    Rectangle (0,0 400x109)
    Rectangle (3,3 394x103), colour toggle: NOT stPis.b_Enable
    Rectangle (209,43 173x61), colour toggle: stPis.st_Open
    Button (220,59 150x30), "%s", text variable: sLable_Open, colour toggle: stPis.req_Open, input disabled if: stPis.b_DeactivateMan OR NOT stPis.b_InterLock_Open
        toggle stPis.req_OpenMan
    RoundedRectangle (260,39 70x15), "open"
    Rectangle (18,43 173x61), colour toggle: stPis.st_Close
    Button (29,59 150x30), "%s", text variable: sLable_Close, colour toggle: stPis.req_Close, input disabled if: stPis.b_DeactivateMan OR NOT stPis.b_InterLock_Close
        toggle stPis.req_CloseMan
    RoundedRectangle (69,39 70x15), "close"
    Button (156,39 83x30), "Default pos", colour toggle: stPis.req_DefaultPos, input disabled if: stPis.b_DeactivateMan
        toggle stPis.req_DefaultPos
    Textfield (5,5 390x33), "piston: %s", text variable: stPis.description
    Textfield (5,7 42x21), "#%d", text variable: stPis.iPisNum
    Button (360,7 35x30), "Err", colour toggle: stPis.b_Error
        toggle stPis.b_Resume
END_VISUALIZATION

// ---- 00 Library/01 Piston/VISU/vis_Piston_Control2_OpenClose.TcVIS
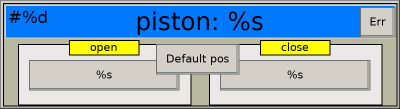
VISUALIZATION vis_Piston_Control2_OpenClose  // 400x109
VAR_IN_OUT
	stPis			: ST_Piston;
END_VAR
VAR_INPUT
	sLable_Open		: STRING:='lable open';
	sLable_Close	: STRING:='lable close';
END_VAR
    Rectangle (0,0 400x109)
    Rectangle (3,3 394x103), colour toggle: NOT stPis.b_Enable
    Rectangle (18,44 173x61), colour toggle: stPis.st_Open
    Rectangle (209,44 173x61), colour toggle: stPis.st_Close
    Button (29,60 150x30), "%s", text variable: sLable_Open, colour toggle: stPis.req_Open, input disabled if: stPis.b_DeactivateMan OR NOT stPis.b_InterLock_Open
        toggle stPis.req_OpenMan
    Button (220,60 150x30), "%s", text variable: sLable_Close, colour toggle: stPis.req_Close, input disabled if: stPis.b_DeactivateMan OR NOT stPis.b_InterLock_Close
        toggle stPis.req_CloseMan
    Button (156,44 83x30), "Default pos", colour toggle: stPis.req_DefaultPos, input disabled if: stPis.b_DeactivateMan
        toggle stPis.req_DefaultPos
    RoundedRectangle (69,40 70x15), "open"
    RoundedRectangle (260,40 70x15), "close"
    Textfield (5,5 390x33), "piston: %s", text variable: stPis.description
    Textfield (5,7 42x21), "#%d", text variable: stPis.iPisNum
    Button (360,7 35x30), "Err", colour toggle: stPis.b_Error
        toggle stPis.b_Resume
END_VISUALIZATION

// ---- 00 Library/01 Piston/VISU/vis_Piston_Select.TcVIS
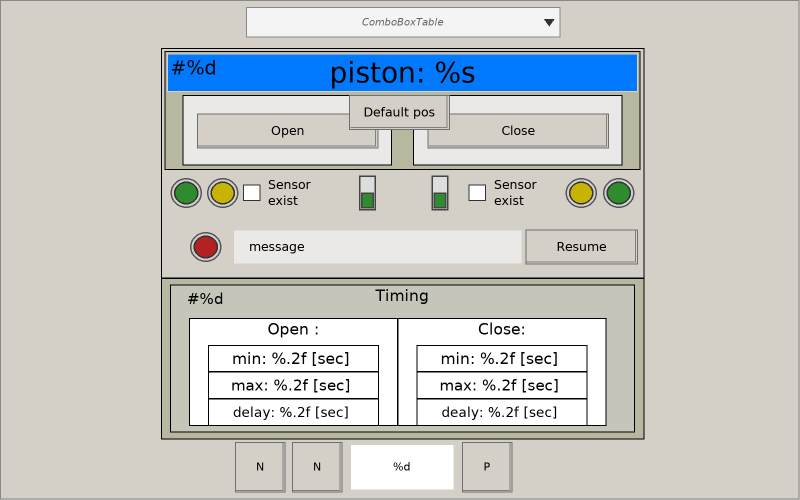
VISUALIZATION vis_Piston_Select  // 800x500
    Frame (161,48 483x230)
        shows vis_Piston_Control1(stPis := stPis[iPis_sel])
    Frame (161,278 483x161)
        shows vis_Piston_Times(stPis := stPis[iPis_sel])
    Button (292,442 50x50), "N"
        tap prg_Piston.bPis_Next_N
    Button (462,442 50x50), "P"
        tap prg_Piston.bPis_Next_P
    Textfield (350,444 104x46), "%d", text variable: iPis_sel
    ComboBoxTable (246,7 314x30), variable: iPis_sel, data array: g_Piston.arPisName
        p3854506369: g_Piston.arPisName[INDEX].Num
        p1892666644: g_Piston.arPisName[INDEX].Description
    Button (235,442 50x50), "N"
        tap prg_Piston.bPis_Next_N
END_VISUALIZATION

// ---- 00 Library/01 Piston/VISU/vis_Piston_Select_1.TcVIS
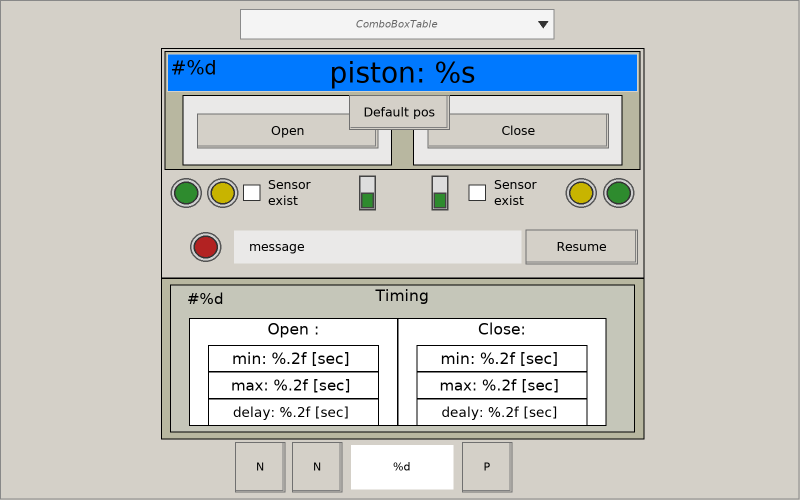
VISUALIZATION vis_Piston_Select_1  // 800x500
    Frame (161,48 483x230)
        shows vis_Piston_Control1(stPis := stPis[iPis_sel])
    Frame (161,278 483x161)
        shows vis_Piston_Times(stPis := stPis[iPis_sel])
    Button (292,442 50x50), "N"
        tap prg_Piston.bPis_Next_N
    Button (462,442 50x50), "P"
        tap prg_Piston.bPis_Next_P
    Textfield (350,444 104x46), "%d", text variable: iPis_sel
    ComboBoxTable (240,9 314x30), variable: iPis_sel, data array: arPisName
        p1128707560: C_MAX_Pistons_Exist
        p3854506369: arPisName[INDEX].Num
        p1892666644: arPisName[INDEX].Description
    Button (235,442 50x50), "N"
        tap prg_Piston.bPis_Next_N
END_VISUALIZATION

// ---- 00 Library/01 Piston/VISU/vis_Piston_Setting_Table.TcVIS
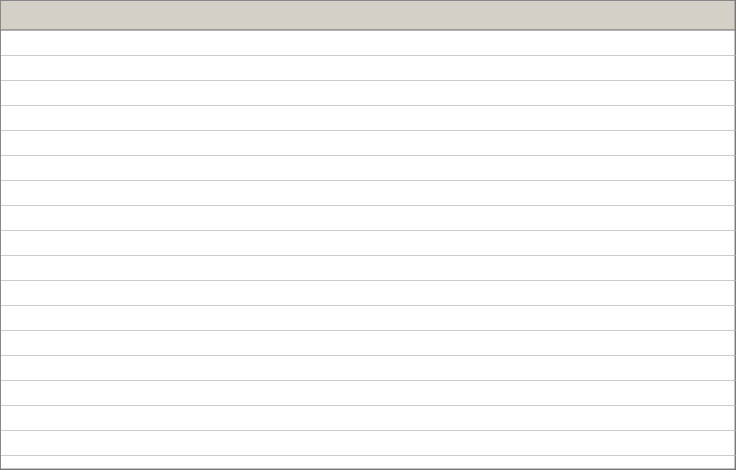
VISUALIZATION vis_Piston_Setting_Table  // 736x470
    Table (0,0 736x470), data array: stPisSetting
        p3854506369: stPisSetting[INDEX].t_minOpen
        p1892666644: stPisSetting[INDEX].t_minClose
        p338671338: stPisSetting[INDEX].t_maxOpen
        p2170511999: stPisSetting[INDEX].t_maxClose
        p3723444502: stPisSetting[INDEX].t_DelayOpen
        p1218418051: stPisSetting[INDEX].t_DelayClose
        p746581629: stPisSetting[INDEX].sen_Open_Exist
        p3104783080: stPisSetting[INDEX].sen_Close_Exist
END_VISUALIZATION

// ---- 00 Library/01 Piston/VISU/vis_Piston_Times.TcVIS
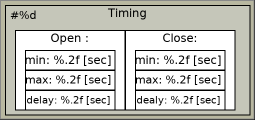
VISUALIZATION vis_Piston_Times  // 255x120
VAR_IN_OUT
	stPis: ST_Piston;
END_VAR
    Rectangle (0,0 255x120)
    Rectangle (5,5 245x110), "Timing"
    Rectangle (15,30 110x80), "Open :"
    Rectangle (125,30 110x80), "Close:"
    Rectangle (135,50 90x20), "min: %.2f [sec]", text variable: stPis.t_minClose
        OnMouseDown: write the text variable via Edit, min 0
    Rectangle (135,70 90x20), "max: %.2f [sec]", text variable: stPis.t_maxClose
        OnMouseDown: write the text variable via Edit, min 0
    Rectangle (25,70 90x20), "max: %.2f [sec]", text variable: stPis.t_maxOpen
        OnMouseDown: write the text variable via Edit, min 0
    Rectangle (25,50 90x20), "min: %.2f [sec]", text variable: stPis.t_minOpen
        OnMouseDown: write the text variable via Edit, min 0
    Rectangle (25,90 90x20), "delay: %.2f [sec]", text variable: stPis.t_DelayOpen
        OnMouseDown: write the text variable via Edit, min 0
    Rectangle (135,90 90x20), "dealy: %.2f [sec]", text variable: stPis.t_DelayClose
        OnMouseDown: write the text variable via Edit, min 0
    Textfield (4,5 39x21), "#%d", text variable: stPis.iPisNum
END_VISUALIZATION

// ---- 00 Library/03 SFC/vis_Cycle_Control.TcVIS
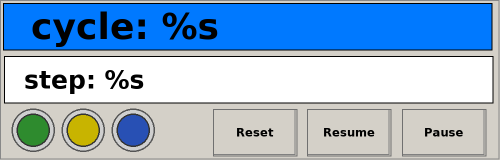
VISUALIZATION vis_Cycle_Control  // 500x160
VAR_IN_OUT
	fb: FB_SFC_Cycle;
END_VAR
VAR_INPUT
	sName: STRING:='Cycle name';
END_VAR
    Lamp1 (8,105 50x50), tooltip "Ready", variable: fb.bReady, style: Lamp-Lamp1-Green
    Lamp1 (108,105 50x50), tooltip "Done", variable: fb.bDone, style: Lamp-Lamp1-Blue
    Lamp1 (58,105 50x50), tooltip "Run", variable: fb.bRun, style: Lamp-Lamp1-Yellow
    RoundedRectangle (3,3 489x47), "cycle: %s", tooltip "POU name: %s", text variable: sName
        p4168582468: fb.refSFC.SFCErrorPOU
    RoundedRectangle (4,56 489x47), "step: %s", text variable: fb.refSFC.SFCCurrentStep, colour toggle: fb.ErrorSFC
    Button (213,109 84x47), "Reset"
        tap fb.bInit
    Button (307,109 84x47), "Resume", colour toggle: fb.ErrorSFC
        toggle fb.refSFC.SFCQuitError
    Button (402,109 84x47), "Pause", colour toggle: fb.refSFC.SFCPause
        toggle fb.refSFC.SFCPause
END_VISUALIZATION

// ---- 00 Library/03 SFC/vis_Cycle_Control_1.TcVIS
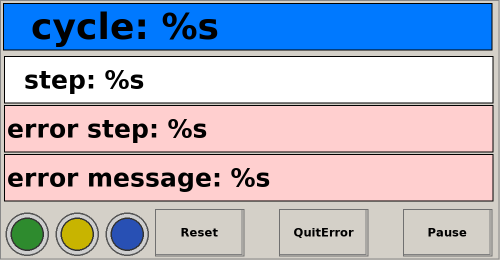
VISUALIZATION vis_Cycle_Control_1  // 500x260
VAR_IN_OUT
	fb: FB_SFC_Cycle;
END_VAR
VAR_INPUT
	sName: STRING:='Cycle name';
END_VAR
    Lamp1 (2,209 50x50), tooltip "Ready", variable: fb.bReady, style: Lamp-Lamp1-Green
    Lamp1 (102,209 50x50), tooltip "Done", variable: fb.bDone, style: Lamp-Lamp1-Blue
    Lamp1 (52,209 50x50), tooltip "Run", variable: fb.bRun, style: Lamp-Lamp1-Yellow
    RoundedRectangle (3,3 489x47), "cycle: %s", tooltip "POU name: %s", text variable: sName
        p4168582468: fb.refSFC.SFCErrorPOU
    RoundedRectangle (4,56 489x47), "step: %s", text variable: fb.refSFC.SFCCurrentStep, colour toggle: fb.ErrorSFC
    Button (155,209 89x47), "Reset"
        tap fb.bInit
    Button (403,209 89x47), "Pause", colour toggle: fb.refSFC.SFCPause
        toggle fb.refSFC.SFCPause
    Button (279,209 89x47), "QuitError", colour toggle: fb.ErrorSFC
        toggle fb.refSFC.SFCQuitError
    RoundedRectangle (4,105 489x47), "error step: %s", text variable: fb.sLastStepBefore_Error, colour toggle: fb.ErrorSFC
    RoundedRectangle (4,154 489x47), "error message: %s", text variable: fb.sError_Message, colour toggle: fb.ErrorSFC
END_VISUALIZATION

// ---- 00 Library/03 SFC/vis_Cycle_Panel.TcVIS
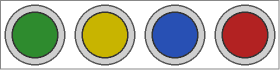
VISUALIZATION vis_Cycle_Panel  // 280x70
VAR_IN_OUT
	fb: FB_SFC_Cycle;
END_VAR
    Lamp1 (0,0 70x70), tooltip "Ready", variable: fb.bReady, style: Lamp-Lamp1-Green
    Lamp1 (70,0 70x70), tooltip "Done", variable: fb.bDone, style: Lamp-Lamp1-Yellow
    Lamp1 (140,0 70x70), tooltip "ToBe Done", variable: fb.bToBe_Done, style: Lamp-Lamp1-Blue
    Lamp1 (210,0 70x70), tooltip "Run", variable: fb.bRun, style: Lamp-Lamp1-Red
END_VISUALIZATION

// ---- 00 Library/04 Recipe/FB_Recipe_Vizu.TcVIS
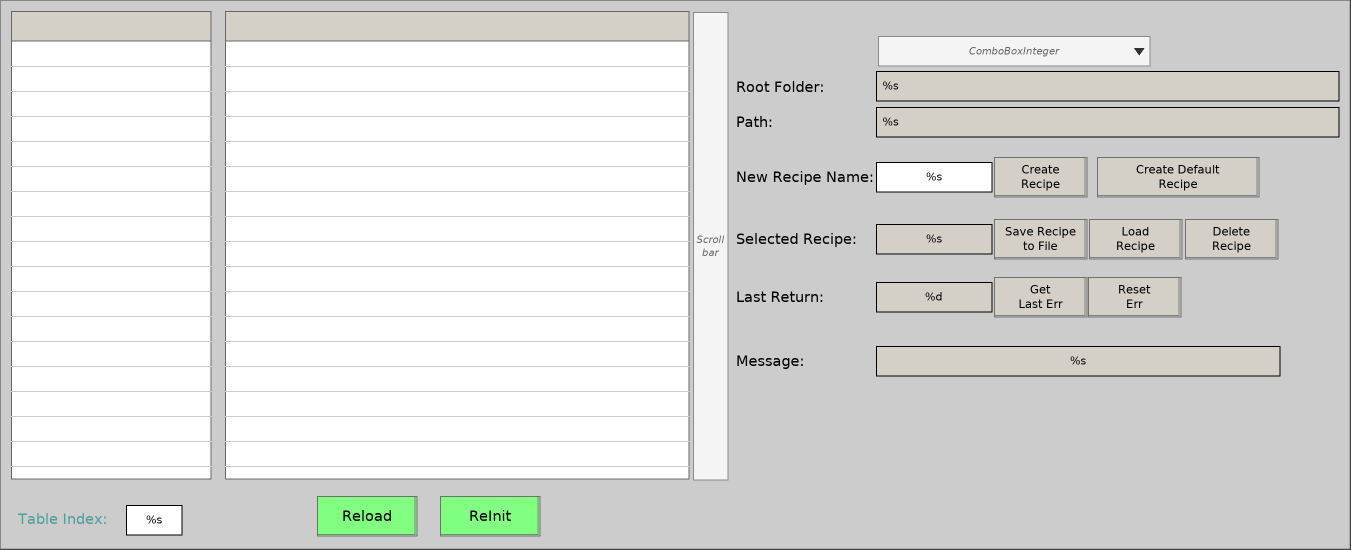
VISUALIZATION FB_Recipe_Vizu  // 1351x550
VAR_IN_OUT
	fb_Recipe		:FB_Recipe;
END_VAR
    Rectangle (0,0 1351x550)
    Table (11,11 200x468), data array: fb_Recipe.pstRecipe^.arrRecipeNames
        p1137915858: fb_Recipe.pstRecipe^.iRecipeIndex
        p1822360349: fb_Recipe.pstRecipe^.bValidSelected
        p3854506369: fb_Recipe.pstRecipe^.arrRecipeNames[INDEX]
        p2232123230: Recipe Names
    Rectangle (126,505 56x30), "%s", text variable: fb_Recipe.pstRecipe^.iRecipeIndex
    Label (15,504 108x30), "Table Index:"
    Button (317,496 100x40), "Reload"
        toggle fb_Recipe.pstRecipe^.bReloadRecipes
    Table (225,11 464x468), data array: fb_Recipe.pstRecipe^.arrVariableDisp
        p3854506369: fb_Recipe.pstRecipe^.arrVariableDisp[0,INDEX]
        p2232123230: No
        p1892666644: fb_Recipe.pstRecipe^.arrVariableDisp[1,INDEX]
        p511219082: Variable Name
        p338671338: fb_Recipe.pstRecipe^.arrVariableDisp[2,INDEX]
        p1755163831: Variable Value
    Scrollbar (693,12 35x468)
        p1057716461: fb_Recipe.pstRecipe^.iDispSel
    Button (1185,219 93x40), "Delete Recipe"
        toggle fb_Recipe.pstRecipe^.bDeleteRecipe
    Label (733,162 141x30), "New Recipe Name:"
    Label (733,224 141x30), "Selected Recipe:"
    Label (733,282 141x30), "Last Return:"
    Rectangle (876,162 116x30), "%s", text variable: fb_Recipe.pstRecipe^.sNewRecipeName
        OnMouseClick: write the text variable via Edit
    Rectangle (876,224 116x30), "%s", text variable: fb_Recipe.pstRecipe^.sSelectedReceipe
    Rectangle (876,282 116x30), "%d", text variable: fb_Recipe.LastReturn, colour toggle: fb_Recipe.LastReturn<>0
    Button (994,157 93x40), "Create Recipe"
        toggle fb_Recipe.pstRecipe^.bCreateRecipe
    Button (994,219 93x40), "Save Recipe to File"
        toggle fb_Recipe.pstRecipe^.bSaveFileCmd
    Button (994,277 93x40), "Get Last Err"
        toggle fb_Recipe.pstRecipe^.bGetLastError
    Button (1089,219 93x40), "Load Recipe"
        toggle fb_Recipe.pstRecipe^.bWriteToPLC_Cmd
    Button (1088,277 93x40), "Reset Err"
        toggle fb_Recipe.pstRecipe^.bResetLastError
    Label (733,107 141x30), "Path:"
    Rectangle (876,107 463x30), "%s", text variable: fb_Recipe.sRecipesStoragePath
    Button (440,496 100x40), "ReInit"
        toggle fb_Recipe.pstRecipe^.bReInit
    Label (733,346 141x30), "Message:"
    Rectangle (876,346 404x30), "%s", text variable: fb_Recipe.sMessage
    Button (1097,157 162x40), "Create Default Recipe"
        toggle fb_Recipe.pstRecipe^.bCreateRecipe
        OnMouseClick: execute { fb_Recipe.pstRecipe^.sNewRecipeName:='Default'; }
    ComboBoxInteger (878,36 272x30), variable: GVL_Recipe.eRecipeRootFolder, text list: 'TextList_RecipeRootFolder'
    Rectangle (876,71 463x30), "%s", text variable: GVL_Recipe.ar_RecipesStoragePath_Root[GVL_Recipe.eRecipeRootFolder]
        OnMouseClick: write the text variable via Edit
    Label (733,72 141x30), "Root Folder:"
END_VISUALIZATION

// ---- 00 Library/04 Recipe/OLD/vis_RecipeControl_v01.TcVIS
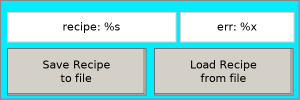
VISUALIZATION vis_RecipeControl_v01  // 300x100
VAR_INPUT
	Definition: STRING;
END_VAR
VAR
	RecipeName: STRING:='name';
END_VAR
    Button (7,48 139x47), "Save Recipe to file"
        OnMouseClick: ExecuteCommand ExecuteCommand=ExecuteCommand=[Command=CreateRecipe, Value=Definition, Value2=RecipeName, Command=SaveRecipeAs, Value=Definition, Value2=RecipeName]
    Button (154,48 139x47), "Load Recipe from file"
        OnMouseClick: ExecuteCommand ExecuteCommand=ExecuteCommand=[Command=LoadRecipeFrom, Value=Definition, Value2=RecipeName]
    Textfield (7,12 169x30), "recipe: %s", text variable: Definition
    Textfield (180,12 114x30), "err: %x", text variable: prg_RecipeManager.LastError, colour toggle: prg_RecipeManager.LastError<>0
        toggle prg_RecipeManager.bResetError
END_VISUALIZATION

// ---- 00 Library/04 Recipe/OLD/vis_RecipeTest.TcVIS
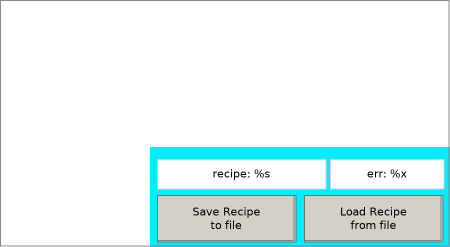
VISUALIZATION vis_RecipeTest  // 450x247
    Frame (150,147 300x100)
        shows vis_RecipeControl_v01(Definition := 'R_Open1')
END_VISUALIZATION

// ---- 00 Library/04 Recipe/TextList_RecipeRootFolder.TcTLO
TEXTLIST TextList_RecipeRootFolder
  0 = 'PLC'
  1 = 'Develop 1'
  2 = 'Develop 2'
  3 = 'Develop 3'
  4 = 'Develop 4'
   = ''
END_TEXTLIST

// ---- 00 Library/05 Safety/Vis_ES_PB.TcVIS
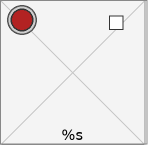
VISUALIZATION Vis_ES_PB  // 148x145
VAR_IN_OUT
	stPB: ST_ES_PB;

END_VAR
VAR_INPUT
	Lable: STRING;

END_VAR
    Image (0,0 145x145), "%s", text variable: Lable, image: ImagePool.EStop_OK2
        p84334746: stPB.stBitMap
    Checkbox (107,3 41x39), tooltip "ByPass", variable: stPB.ByPass, input disabled if: prg_User.actUser<4
    Lamp1 (5,3 34x34), tooltip "Memo PB State", variable: stPB.Memo, style: Lamp-Lamp1-Red
END_VISUALIZATION

// ---- 00 Library/06-Visu/Sensor.TcVIS
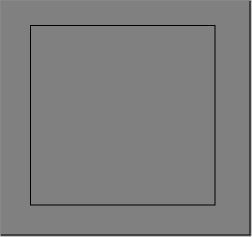
VISUALIZATION Sensor  // 252x237
VAR_INPUT
	{attribute 'parameterstringof' := 'm_Input_Sen_Addr'}
	m_Input_Sen_Addr_Str : STRING;
END_VAR
VAR_INPUT
	m_Input_Sen_Addr : Bool;
END_VAR
    Rectangle (0,0 250x235)
    RoundedRectangle (30,25 185x180), tooltip "%s", colour toggle: (m_Input_Sen_Addr) <> 0
        p4168582468: m_Input_Sen_Addr_Str
END_VISUALIZATION

// ---- 00 Library/07 Errors/vis_Device_Error.TcVIS
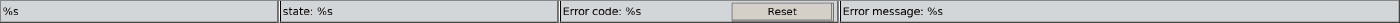
VISUALIZATION vis_Device_Error  // 1500x25
VAR_IN_OUT
	fb_comm_dev: fb_common_device;
END_VAR
    Rectangle (900,0 600x25), "Error message: %s", text variable: fb_comm_dev.common_events.device_error.error_string, colour toggle: fb_comm_dev.common_events.device_error.error_code<>''
        OnMouseUp: execute { GVL.Errors:=(0); }
    Rectangle (600,0 298x25), "Error code: %s", text variable: fb_comm_dev.common_events.device_error.error_code, colour toggle: fb_comm_dev.common_events.device_error.error_code<>''
        OnMouseUp: execute { GVL.Errors:=(0); }
    Button (784,3 109x20), "Reset"
        toggle fb_comm_dev.common_actions.reset
    Rectangle (0,0 298x25), "%s", tooltip "Device Name", text variable: fb_comm_dev.Name, colour toggle: fb_comm_dev.common_events.device_error.error_code<>''
        OnMouseUp: execute { GVL.Errors:=(0); }
    Rectangle (300,0 298x25), "state: %s", tooltip "Device State", text variable: fb_comm_dev.device_status, colour toggle: fb_comm_dev.common_events.device_error.error_code<>''
        OnMouseUp: execute { GVL.Errors:=(0); }
END_VISUALIZATION

// ---- 00 Library/07-Mode/Visu/Mode_Select.TcVIS
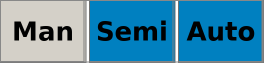
VISUALIZATION Mode_Select  // 264x63
VAR_IN_OUT
	stMode: ST_Mode;
END_VAR
    Button (0,0 86x63), "Man", colour toggle: stModeMain.iActMode=eManualMode
        OnMouseDown: execute {
            stModeMain.bSetManual:=TRUE;
            stMode.bSetSemi:=FALSE;
            stMode.bSetAuto:=FALSE;
        }
    Button (89,0 86x63), "Semi", colour toggle: stModeMain.iActMode=eSemiAutoMode
        OnMouseDown: execute {
            stModeMain.bSetManual:=FALSE;
            stMode.bSetSemi:=TRUE;
            stMode.bSetAuto:=FALSE;
        }
    Button (178,0 86x63), "Auto", colour toggle: stModeMain.iActMode=eAutoMode
        OnMouseDown: execute {
            stModeMain.bSetManual:=FALSE;
            stMode.bSetSemi:=FALSE;
            stMode.bSetAuto:=TRUE;
        }
END_VISUALIZATION

// ---- 00 Library/07-Mode/Visu/Mode_Select_1.TcVIS
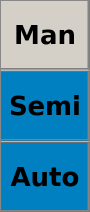
VISUALIZATION Mode_Select_1  // 90x212
VAR_IN_OUT
	stMode: ST_Mode;
END_VAR
    Button (0,0 90x70), "Man", colour toggle: stModeMain.iActMode=eManualMode, input disabled if: NOT GVL.MainMachine.bReadyToManualModeSelect
        OnMouseDown: execute {
            stModeMain.bSetManual:=TRUE;
            stMode.bSetSemi:=FALSE;
            stMode.bSetAuto:=FALSE;
        }
    Button (0,71 90x70), "Semi", colour toggle: stModeMain.iActMode=eSemiAutoMode, input disabled if: stModeMain.iActMode<>E_WorkingMode.eManualMode
        OnMouseDown: execute {
            stModeMain.bSetManual:=FALSE;
            stMode.bSetSemi:=TRUE;
            stMode.bSetAuto:=FALSE;
        }
    Button (0,142 90x70), "Auto", colour toggle: stModeMain.iActMode=eAutoMode, input disabled if: stModeMain.iActMode<>E_WorkingMode.eManualMode
        OnMouseDown: execute {
            stModeMain.bSetManual:=FALSE;
            stMode.bSetSemi:=FALSE;
            stMode.bSetAuto:=TRUE;
        }
END_VISUALIZATION

// ---- 00 Library/07-Mode/Visu/OperationButtons.TcVIS
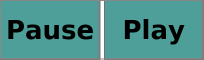
VISUALIZATION OperationButtons  // 204x60
VAR_IN_OUT
	stOperation	:ST_OperationButtons;
END_VAR
    Button (0,0 100x60), "Pause", tooltip "%s", colour toggle: stOperation.iActOperation=ePauseAll
        p4168582468: stOperation.sModeZone
        OnMouseClick: execute { stOperation.bSetPause:=TRUE; stOperation.iPauseHistory:=7; }
    Button (104,0 100x60), "Play", tooltip "%s", colour toggle: stOperation.iActOperation=ePlayAll
        p4168582468: stOperation.sModeZone
        OnMouseClick: execute { stOperation.bSetPlay:=TRUE; }
END_VISUALIZATION

// ---- 00 Library/07-Mode/Visu/OperationButtons_1.TcVIS
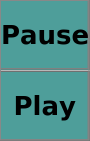
VISUALIZATION OperationButtons_1  // 90x141
VAR_IN_OUT
	stOperation	:ST_OperationButtons;
END_VAR
    Button (0,0 90x70), "Pause", colour toggle: stOperation.iActOperation=ePauseAll
        OnMouseClick: execute { stOperation.bSetPause:=TRUE; stOperation.iPauseHistory:=7; }
    Button (0,71 90x70), "Play", colour toggle: stOperation.iActOperation=ePlayAll
        OnMouseClick: execute { stOperation.bSetPlay:=TRUE; }
END_VISUALIZATION

// ---- 00 Library/07-Mode/Visu/OperationButton_Stop.TcVIS
